(* IEC 61131-3 sources: daoli-st-library/DL_Motion (part 15) *)

(* ---- FB_DL_LaserTabWeldTrack.st ---- *)
(*==============================================================================
 * 组件名称 (Component)  : FB_DL_LaserTabWeldTrack
 * 所属子库 (Sublibrary) : DL_Motion
 * 当前版本 (Version)    : 1.0.1
 * 兼容性 (Platform)     : CODESYS 3.5 / TwinCAT 3 / 汇川 InoProShop（纯标准元素，零方言）
 * 功能描述 (Function)   : 极耳激光焊跟随误差与虚焊特征窗监视。出光期间统计三类缺陷特征
 *                         ——跟随误差超限、功率相对跌落、位置停滞——各需连续满足确认时长
 *                         才置位；单焊点窗口超时强制给出判决并置超时位，绝不允许无限期停
 *                         在出光态。不做激光功率闭环、不做焊缝跟踪插补、不做焊后强度判定。
 *                         交付门槛：位置停滞判据用 tConfirm 换算秒（时间转换链），须在
 *                         CODESYS / TwinCAT / InoProShop 三平台各编译验证一次。
 * 溯源 (Origin)         : 道莅 clean-room 防御性实现
 * 本文件内含 (Contains) : TYPE E_DL_WeldTrackState / FUNCTION_BLOCK FB_DL_LaserTabWeldTrack
 * 依赖 (Depends)        : 无（仅 Standard.library 的 ABS / MAX / TIME_TO_LREAL）
 * 红线自检 (Redline)    : 无外部全局变量、无硬件地址直引 ｜ 全变量中英双语同行注释
 *                         参考功率与误差上限判零防除零 ｜ 位置非有限只跳过本拍、不清峰值
 *                         四个定时器无条件周期刷新 ｜ 枚举显式赋值 ｜ CASE 含 ELSE 兜底
 * 同拍双窗配比约束      : 窗口超时 tWindowMax 必须显著大于三类判据确认 tConfirm
 *                         （建议 tWindowMax ≥ 5 × tConfirm），否则判据来不及确认即被超时
 *                         抢先判决，缺陷掩码永远只能出 bit3。
 * 错误码表 (Codes)      : 16#0004_0331 就绪（无窗进行或本拍无故障）
 *                         16#0004_0332 信息级 位置读数非有限，本拍跳过（已累计峰值与掩码
 *                                    保持，不清零）
 *                         16#0004_0333 故障级 组态非法（跟随误差上限或参考功率 ≤0）
 *                         16#0004_0334 故障级 非法状态兜底（状态机落 ELSE）
 *                         16#0004_0335 预留：本版不发码（下一轮区间起点，禁止回填）
 * 修订历史 (Revision)   : 2026-11-17  v1.0.0  首版入库 · R28 · 阶段三批 2
 *                         2026-11-17  v1.0.1  终审修复：①停滞速度补入组态域闸（负值/NaN 会
 *                                    使停滞距离门限失效而静默关闭 bit2 判据）；②停滞窗起点与
 *                                    焊点位置锁存加位置有限前置（防 NaN 写入出口）· R28 · 阶段四
 * 验收向量 (Acceptance) : 正向 指令 0→50 mm、实际滞后 0.3 mm 超上限 0.2 mm 持续 30 ms →
 *                         bit0 置位、eState=eReject、峰值 0.3 mm
 *                         反向 功率 2000→1500 W（跌 25% 超 10%）持续 30 ms → bit1；
 *                         上限给 0 → 16#0004_0333；窗口拖满 tWindowMax 无判决 → bit3 +
 *                         eReject（不停在出光态）；位置给 NaN → 16#0004_0332 且峰值不清零
 *============================================================================*)

(*-----------------------------------------------------------------------------
 * 枚举: E_DL_WeldTrackState（归属本功能块，同文件发布，全库唯一定义）
 * 含义: 单焊点监视相位，每个成员在 CASE 中有且仅有一个标签。
 *----------------------------------------------------------------------------*)
TYPE E_DL_WeldTrackState :
(
    eWaiting  := 0,    // 待机：等出光 / Waiting for the weld-on signal
    eWelding  := 10,   // 出光中：累计峰值与三类判据 / Welding, accumulating the peak and the three criteria
    eJudging  := 20,   // 判决中：锁存焊点位置并出结论 / Judging, latching the weld position and issuing the verdict
    ePass     := 30,   // 合格：掩码为 0 / Pass, the defect mask is zero
    eReject   := 40,   // 不合格：至少一个缺陷位或窗口超时 / Reject, at least one defect bit or the window timed out
    eFault    := 99    // 故障：锁存码保持，仅使能沿重启 / Fault, the latch code is held until an enable edge
);
END_TYPE

FUNCTION_BLOCK FB_DL_LaserTabWeldTrack
VAR_INPUT
    bEnable         : BOOL := FALSE;      // 使能 / Enable
    bWeldOn         : BOOL := FALSE;      // 出光中（仅窗内判据） / Welding on, the criteria are evaluated inside the window only
    fPosCmd_mm      : REAL := 0.0;        // 指令位置 [mm] / Command position in millimetres
    fPosAct_mm      : REAL := 0.0;        // 实际位置 [mm] / Actual position in millimetres
    fPower_W        : REAL := 0.0;        // 实测功率 [W] / Measured power in watt
    fPowerRef_W     : REAL := 2000.0;     // 设定功率 [W]，须 >0 / Reference power in watt, must be positive
    fFollowErrMax_mm : REAL := 0.2;       // 跟随误差上限 [mm]，域 0.01~2.0 / Following error limit in millimetres, domain 0.01 to 2.0
    fPowerDropPct   : REAL := 10.0;       // 功率跌落阈 [%]，域 1~50 / Power drop threshold in percent, domain 1 to 50
    fStallVel_mmS   : REAL := 0.2;        // 停滞判据速度 [mm/s]，域 0~5 / Stall speed criterion in millimetres per second, domain 0 to 5
    tConfirm        : TIME := T#30MS;     // 判据确认时长 [ms]，域 20~500 / Criterion confirmation time, domain 20 to 500 ms
    tWindowMax      : TIME := T#2S;       // 单焊点窗口 [ms]，域 50ms~10s / Single weld spot window, domain 50 ms to 10 s
END_VAR
VAR_OUTPUT
    bTrackOk        : BOOL;               // 轨迹合格（判决合格时置位） / Trajectory accepted
    fFollowErrPeak_mm : REAL;             // 窗内跟随误差峰值 [mm] / Peak following error inside the window
    uDefectMask     : WORD;               // 缺陷掩码 bit0 跟超 bit1 功率跌 bit2 停滞 bit3 超时 [bit] / Defect mask
    fWeldPos_mm     : REAL;               // 锁存焊点位置 [mm] / Latched weld position in millimetres
    eState          : E_DL_WeldTrackState; // 监视相位 [—] / Monitoring phase
    eErr            : UDINT;              // 错误码，段位 16#0004_xxxx / Error code in segment 16#0004_xxxx
END_VAR
VAR
    _eState         : E_DL_WeldTrackState := E_DL_WeldTrackState.eWaiting; // 当前相位 / Current phase
    _bInit          : BOOL := FALSE;      // 首扫标志，取非判定 / First-scan flag, tested negated
    _bCfgOk         : BOOL;               // 组态合法标志 / Configuration valid flag
    _bPosOk         : BOOL;               // 位置读数有限标志 / Position readings finite flag
    _bFaultLatch    : BOOL;               // 故障锁存标志 / Fault latch flag
    _uLatchCode     : UDINT;              // 锁存码载体 / Latch code carrier
    _fFollowErr     : REAL;               // 本拍跟随误差 [mm] / Following error of this scan
    _fPeak          : REAL;               // 窗内峰值内部副本 [mm] / Internal peak copy inside the window
    _fDropPct       : REAL;               // 本拍功率跌落百分比 [%] / Power drop of this scan in percent
    _fPosWinStart   : REAL;               // 停滞窗起点位置 [mm] / Position at the start of the stall window
    _fConfirmSec    : REAL := 0.03;       // 确认时长换算秒 [s] / Confirmation time converted to seconds
    _fStallDist     : REAL;               // 停滞判定距离门限 [mm] / Stall distance threshold in millimetres
    _rtrigEnable    : R_TRIG;             // 使能上升沿 / Rising edge of the enable input
    _tonFollow      : TON;                // 跟超确认计时 / Following error confirmation timer
    _tonPower       : TON;                // 功率跌落确认计时 / Power drop confirmation timer
    _tonStall       : TON;                // 停滞确认计时 / Stall confirmation timer
    _tonWindow      : TON;                // 单焊点窗口计时 / Weld spot window timer
END_VAR
VAR CONSTANT
    DL_WT_READY     : UDINT := 16#0004_0331;  // 就绪码 / Ready code
    DL_WT_POS_BAD   : UDINT := 16#0004_0332;  // 信息级位置非有限码 / Info code for non-finite positions
    DL_WT_CFG_BAD   : UDINT := 16#0004_0333;  // 故障级组态非法码 / Fault code for bad configuration
    DL_WT_ILLEGAL   : UDINT := 16#0004_0334;  // 故障级非法状态码 / Fault code for an illegal state
    DL_WT_BIT_FOLLOW : WORD := 16#0001;       // 缺陷位 bit0 跟超 / Defect bit 0, following error
    DL_WT_BIT_POWER  : WORD := 16#0002;       // 缺陷位 bit1 功率跌 / Defect bit 1, power drop
    DL_WT_BIT_STALL  : WORD := 16#0004;       // 缺陷位 bit2 停滞 / Defect bit 2, stall
    DL_WT_BIT_TIME   : WORD := 16#0008;       // 缺陷位 bit3 超时 / Defect bit 3, window timeout
    DL_WT_EPS        : REAL := 1.0E-6;        // 浮点判零容差 [—] / Float zero tolerance
END_VAR

// 段 1｜输出与单拍标志预置（bTrackOk 逐拍重算，掩码与峰值为窗内累计量，不在此清）
bTrackOk := FALSE;                                  // 合格标志预清 / Accepted flag pre-cleared
eErr := 0;                                          // 错误码预清 / Error code pre-cleared

// 段 2｜沿检测无条件周期刷新
_rtrigEnable(CLK := bEnable);                       // 使能沿 / Enable edge

// 段 3｜首扫初始化（判据取非，R19）
IF NOT _bInit THEN
    _eState := E_DL_WeldTrackState.eWaiting;        // 相位待机起步 / Phase starts waiting
    _bInit := TRUE;                                 // 首扫只做一次 / The first scan runs once
END_IF

// 段 4｜组态闸（跟随上限与参考功率判零防除零）
_bCfgOk := NOT ((fFollowErrMax_mm <> fFollowErrMax_mm) OR ((fFollowErrMax_mm - fFollowErrMax_mm) <> (fFollowErrMax_mm - fFollowErrMax_mm)))
        AND (fFollowErrMax_mm > DL_WT_EPS)
        AND NOT ((fPowerRef_W <> fPowerRef_W) OR ((fPowerRef_W - fPowerRef_W) <> (fPowerRef_W - fPowerRef_W)))
        AND (fPowerRef_W > DL_WT_EPS)
        AND (fPowerDropPct >= 1.0) AND (fPowerDropPct <= 50.0)
        AND (fStallVel_mmS >= 0.0) AND (fStallVel_mmS <= 5.0)   // 停滞速度域闸：负值/NaN 会使停滞门限失效而静默关闭 bit2 / Stall speed gate, a negative or NaN value silently disables bit 2
        AND (tConfirm >= T#20MS) AND (tConfirm <= T#500MS)
        AND (tWindowMax >= T#50MS) AND (tWindowMax <= T#10S);
_fConfirmSec := TIME_TO_LREAL(tConfirm) / 1000.0;   // 确认时长换算秒 [s] / Confirmation time in seconds
_fStallDist := fStallVel_mmS * _fConfirmSec;        // 停滞判定距离门限 [mm] / Stall distance threshold

// 段 5｜位置有限闸（非有限只跳过本拍，已累计峰值与掩码一律不清零）
_bPosOk := NOT ((fPosCmd_mm <> fPosCmd_mm) OR ((fPosCmd_mm - fPosCmd_mm) <> (fPosCmd_mm - fPosCmd_mm)))
        AND NOT ((fPosAct_mm <> fPosAct_mm) OR ((fPosAct_mm - fPosAct_mm) <> (fPosAct_mm - fPosAct_mm)));
_fFollowErr := ABS(fPosCmd_mm - fPosAct_mm);        // 本拍跟随误差 [mm] / Following error of this scan

// 段 6｜功率跌落百分比（除数已在段 4 判零）
IF (fPower_W <> fPower_W) OR ((fPower_W - fPower_W) <> (fPower_W - fPower_W)) THEN
    _fDropPct := 0.0;                               // 功率非有限：本拍不判跌落 / Non-finite power, no drop judgement this scan
ELSE
    _fDropPct := ((fPowerRef_W - fPower_W) / fPowerRef_W) * 100.0;   // 跌落百分比 [%] / Power drop in percent
END_IF

// 段 7｜四个定时器无条件周期刷新（严禁置于分支内）
_tonFollow(IN := (_eState = E_DL_WeldTrackState.eWelding) AND _bPosOk AND (_fFollowErr > fFollowErrMax_mm), PT := tConfirm);
_tonPower(IN := (_eState = E_DL_WeldTrackState.eWelding) AND (_fDropPct > fPowerDropPct), PT := tConfirm);
_tonStall(IN := (_eState = E_DL_WeldTrackState.eWelding) AND _bPosOk AND (ABS(fPosAct_mm - _fPosWinStart) < _fStallDist), PT := tConfirm);
_tonWindow(IN := (_eState = E_DL_WeldTrackState.eWelding), PT := tWindowMax);

// 段 8｜使能上升沿：锁存解除路径
IF _rtrigEnable.Q THEN
    _bFaultLatch := FALSE;                          // 锁存解除 / Latch released
    _uLatchCode := 0;                               // 锁存码清 / Latch code cleared
    _eState := E_DL_WeldTrackState.eWaiting;        // 相位回待机 / Phase back to waiting
    uDefectMask := 16#0000;                         // 掩码清 / Defect mask cleared
    _fPeak := 0.0;                                  // 峰值清 [mm] / Peak cleared
    fFollowErrPeak_mm := 0.0;                       // 峰值出口清 [mm] / Peak output cleared
END_IF

// 段 9｜失能闸
IF NOT bEnable THEN
    _eState := E_DL_WeldTrackState.eWaiting;        // 相位回待机 / Phase back to waiting
    eErr := DL_WT_READY;                            // 失能为正常停机 / Disable is a normal stop
END_IF

// 段 10｜监视状态机（ENUM + CASE + ELSE 兜底）
IF bEnable THEN
    CASE _eState OF

        E_DL_WeldTrackState.eWaiting:               // 待机：组态错即锁存，出光沿开窗
            IF NOT _bCfgOk THEN
                eErr := DL_WT_CFG_BAD;              // 故障级：组态非法 / Fault, bad configuration
                _uLatchCode := DL_WT_CFG_BAD;
                _bFaultLatch := TRUE;
                _eState := E_DL_WeldTrackState.eFault;
            ELSIF bWeldOn THEN
                uDefectMask := 16#0000;             // 新焊点掩码清 / New spot, the mask is cleared
                _fPeak := 0.0;                      // 新焊点峰值清 [mm] / New spot, the peak is cleared
                fFollowErrPeak_mm := 0.0;
                IF _bPosOk THEN                     // 位置有限才取窗起点与焊点初值（防 NaN 入出口） / Latch only with finite positions
                    _fPosWinStart := fPosAct_mm;    // 停滞窗起点位置 [mm] / Stall window start position
                    fWeldPos_mm := fPosAct_mm;      // 焊点位置初值 [mm] / Weld position initial value
                END_IF
                _eState := E_DL_WeldTrackState.eWelding;   // 开窗出光 / The window opens
            ELSE
                eErr := DL_WT_READY;                // 就绪码 / Ready code
            END_IF

        E_DL_WeldTrackState.eWelding:               // 出光中：累计峰值 + 三类判据确认
            IF NOT _bPosOk THEN
                eErr := DL_WT_POS_BAD;              // 信息级：位置非有限，本拍跳过 / Info, positions not finite, this scan is skipped
            ELSE
                IF _fFollowErr > _fPeak THEN
                    _fPeak := _fFollowErr;          // 峰值刷新 [mm] / Peak refreshed
                END_IF
            END_IF
            fFollowErrPeak_mm := _fPeak;            // 峰值出口 [mm] / Peak output
            IF _fFollowErr > fFollowErrMax_mm THEN
                IF _tonFollow.Q THEN
                    uDefectMask := uDefectMask OR DL_WT_BIT_FOLLOW;   // bit0 跟超确认 / Following error confirmed
                END_IF
            END_IF
            IF _fDropPct > fPowerDropPct THEN
                IF _tonPower.Q THEN
                    uDefectMask := uDefectMask OR DL_WT_BIT_POWER;    // bit1 功率跌落确认 / Power drop confirmed
                END_IF
            END_IF
            IF ABS(fPosAct_mm - _fPosWinStart) < _fStallDist THEN
                IF _tonStall.Q THEN
                    uDefectMask := uDefectMask OR DL_WT_BIT_STALL;    // bit2 停滞确认 / Stall confirmed
                END_IF
            ELSE
                _fPosWinStart := fPosAct_mm;    // 已移动：重置停滞窗起点 [mm] / Moved, restart the stall window
            END_IF
            IF _tonWindow.Q THEN
                uDefectMask := uDefectMask OR DL_WT_BIT_TIME;         // bit3 窗口超时 / Window timed out
                _eState := E_DL_WeldTrackState.eJudging;              // 强制判决，绝不停在出光态 / Forced verdict, never stuck in welding
            ELSIF NOT bWeldOn THEN
                _eState := E_DL_WeldTrackState.eJudging;              // 出光结束：判决 / Weld finished, judge now
            END_IF

        E_DL_WeldTrackState.eJudging:               // 判决中：锁存焊点位置并出结论
            IF _bPosOk THEN                         // 位置有限才刷新焊点位置，保持上次有效值 / Refresh the latch only with finite positions
                fWeldPos_mm := fPosAct_mm;          // 锁存焊点位置 [mm] / Latch the weld position
            END_IF
            IF uDefectMask = 16#0000 THEN
                bTrackOk := TRUE;                   // 掩码为 0：合格 / A zero mask means pass
                _eState := E_DL_WeldTrackState.ePass;
            ELSE
                _eState := E_DL_WeldTrackState.eReject;   // 有缺陷位：不合格 / At least one defect bit, reject
            END_IF
            eErr := DL_WT_READY;                    // 判决本身无故障码 / The verdict produces no fault code

        E_DL_WeldTrackState.ePass:                  // 合格：保持结论，等出光消失后回待机
            bTrackOk := TRUE;
            IF NOT bWeldOn THEN
                _eState := E_DL_WeldTrackState.eWaiting;
            END_IF

        E_DL_WeldTrackState.eReject:                // 不合格：保持结论，等出光消失后回待机
            bTrackOk := FALSE;
            IF NOT bWeldOn THEN
                _eState := E_DL_WeldTrackState.eWaiting;
            END_IF

        E_DL_WeldTrackState.eFault:                 // 故障：锁存码保持
            eErr := _uLatchCode;                    // 锁存码回放 / Replay the latch code
            IF NOT _bFaultLatch THEN
                _eState := E_DL_WeldTrackState.eWaiting;   // 锁存已由使能沿解除 / The latch was released by the enable edge
            END_IF

        ELSE
            // 非法状态兜底（故障级）
            eErr := DL_WT_ILLEGAL;                  // 故障级：非法相位 / Fault, illegal phase
            _uLatchCode := DL_WT_ILLEGAL;
            _bFaultLatch := TRUE;
            _eState := E_DL_WeldTrackState.eFault;

    END_CASE
END_IF

eState := _eState;                                  // 相位出口镜像 / Phase mirrored to the output pin
END_FUNCTION_BLOCK

(* ---- FB_DL_LineShaftClutch.st ---- *)
(*
  FB_DL_LineShaftClutch  —  线轴电子离合器（相位对齐 / 咬合 / 打滑监视 / 强制脱开）/ Line-shaft electronic clutch
  分类 Category : DL_Motion
  码位 Code     : 16#04_0_A2
  版本 Version  : 1.0.2
  来源 Source   : t2-4-s7-motion — IEC 61131-3 标准语义的道莅防御性实现
  溯源 Origin   : S7 Motion Control 公开语义借鉴（电子离合器 / 相位偏移 / 打滑监视），clean-room 实现，未复制源码行
  功能 Function : 1) 对齐段：按相位误差（从轴位置 − 主轴位置 − fPhaseOffsetDeg，归一化到 ±180°）输出修正速度
                     指令 fTrimVelDegS，供下游电子齿轮/速度环消费，误差进 fAlignTolDeg（本件常量 0.5°）后进咬合；
                  2) 咬合段：按 fEngageRampTime 斜坡把同步权重从 0 升到 1，斜坡溢出（TON.Q）置 bEngaged；
                     脱开权重自进入脱开相的实际权重按斜坡线性回落到 0，禁跳变到满值（R38 返修口径）；
                  3) 咬合期监视相位误差，超 fSlipLimitDeg 持续 tSlipDebounce → bSlipFault 锁存并强制脱开；
                  4) 脱开段：按同一斜坡时间把同步权重降回 0，权重回零才回 eIdle（不留残余同步量）。
  边界 Boundary : ① fEngageRampTime <= 0 或 fSlipLimitDeg <= 0 判组态错置 00A2，状态进 eFault 不投运；
                  ② 两轴任一 bError / 非 bEnabled → 拒绝咬合并置信息级 05A2（不置 bError，故障属主是轴本身）；
                  ③ 主从同轴（同一实例注入两侧）判组态错置 04A2：接口契约无指针恒等比较（R28 禁臆造），
                     本件改用**代理判据**——连续 DL_SAME_CYC 拍内两轴位置与速度差均 < 1E-6 且至少一侧使能，
                     视为同一实例注入（说明见「同轴代理判据」段）；
                  ④ 脱开命令与咬合命令同拍 → 以脱开为安全优先（脱开优先判定在本段最前），并置 02A2；
                  ⑤ 咬合中主轴反转（速度 < 0）判工装条件越界 → 强制脱开并置 03A2（反转咬合会拉断机械）；
                  ⑥ bSlipFault 解除式 = bReset AND 主轴 eState = eStandstill AND 从轴 eState = eStandstill
                     （三条件均由注入轴的 PROPERTY 可读，R28-1 通过；接口无 bStandstill 属性，改用
                     E_DL_AxisState.eStandstill 判等，属契约内等价表达，已在头注释声明）。
  依赖 Depends  : I_DL_MotionAxis / E_DL_AxisState（DL_Motion 既有契约件，零修改，仅注入不实例化）；
                  仅 Standard.library（TON / R_TRIG / ABS / MAX / MIN）
  同拍双窗配比  : tSlipDebounce（打滑去抖窗）与 fEngageRampTime 不同源；配比约束
                  tSlipDebounce <= fEngageRampTime × 1000 ms，避免咬合斜坡未完成就打滑判据成立（R100）

  码表 Error codes（本件格 04_0_A2，子码步进 +0x10）:
    16#0004_00A2 故障级：组态非法（斜坡时间 <= 0 / 打滑门限 <= 0 / 对齐容差 <= 0）
    16#0004_01A2 故障级：打滑故障锁存（相位误差超 fSlipLimitDeg 持续 tSlipDebounce，已强制脱开）
    16#0004_02A2 故障级：咬合与脱开命令同拍冲突（脱开优先执行，本码锁存待复位确认）
    16#0004_03A2 故障级：咬合期主轴反转（工装条件越界，已强制脱开）
    16#0004_04A2 故障级：主从同轴注入（代理判据成立，组态错）
    16#0004_05A2 信息级：拒绝咬合（注入轴故障或未使能，不置 bError）
    16#0004_06A2 信息级：咬合完成（bEngaged 上升拍，不置 bError）
    16#0004_07A2 故障级：状态机落 ELSE 兜底（非法相位 ID）
    16#0004_08A2 信息级：脱开起始权重为 0，单拍收口（R38 返修新增，不置 bError）

  修订历史 Revision :
    2026-11-18  v1.0.0  R37 首版
    2026-11-18  v1.0.2  R38 返修：脱离相权重起始值改为进入脱开相快照按斜坡线性回落（_fW0Diseng），起始权重 0 单拍收口，消除反向驱动风险
  R38 已修复    : R37 终审挂账「脱离相耦合权重起始值取成满值」已按快照回落方案修复（六处置相点全部先快照后置相）
*)

TYPE E_DL_ClutchState :
(
    eIdle        := 0,   // 空闲：同步权重 0，等待咬合命令 / Idle, sync weight zero
    eAligning    := 10,  // 对齐中：相位误差收敛至容差内 / Aligning, phase error inside the tolerance
    eRamping     := 20,  // 咬合斜坡中：同步权重 0→1 / Engage ramp, weight rising from zero to one
    eEngaged     := 30,  // 已咬合：同步权重 1，监视打滑 / Engaged, weight one, slip supervised
    eDisengaging := 40,  // 脱开斜坡中：同步权重 1→0 / Disengage ramp, weight falling to zero
    eFault       := 50   // 故障：锁存待复位（复位且两轴静止）/ Fault, latched until reset with both axes standstill
);
END_TYPE

FUNCTION_BLOCK FB_DL_LineShaftClutch
VAR_INPUT
    bEnable        : BOOL := FALSE;              // 总使能，FALSE 时按脱开处理 / Master enable, a low level disengages
    bReset         : BOOL := FALSE;              // 复位，上升沿清故障锁存（须两轴静止）/ Reset, clears the latch when both axes stand still
    bEngageCmd     : BOOL := FALSE;              // 咬合命令（电平，保持型）/ Engage command, level held by the caller
    bDisengageCmd  : BOOL := FALSE;              // 脱开命令（电平，安全优先）/ Disengage command, safety priority
    fPhaseOffsetDeg : REAL := 0.0;               // 从轴相对主轴的相位偏移 [°]，域 ±360 / Phase offset of the slave relative to the master [deg]
    fEngageRampTime : REAL := 0.5;               // 咬合/脱开斜坡时间 [s]，域 > 0 / Engage and disengage ramp time [s]
    fSlipLimitDeg  : REAL := 2.0;                // 打滑门限（相位误差绝对值）[°]，域 > 0 / Slip limit [deg]
    tSlipDebounce  : TIME := T#200MS;            // 打滑去抖窗 [ms]，域 > 0 / Slip debounce window [ms]
    fSlipReleaseBandDeg : REAL := 0.2;           // 打滑解除带回差 [°]，域 >= 0 / Slip release hysteresis band [deg]
END_VAR
VAR_OUTPUT
    bEngaged       : BOOL;                       // 已咬合标志（同步权重达 1）/ Engaged flag, sync weight reached one
    bSlipFault     : BOOL;                       // 打滑故障锁存出口 / Slip fault latch outlet
    fPhaseErrorDeg : REAL;                       // 归一化相位误差 [°]，域 ±180 / Normalised phase error [deg]
    fTrimVelDegS   : REAL;                       // 对齐修正速度指令 [°/s]，带符号 / Alignment trim velocity command [deg/s]
    fSyncWeight    : REAL;                       // 同步权重 [0~1]，供下游齿轮/速度环 / Sync weight for the downstream gear or velocity loop
    bAxesReady     : BOOL;                       // 两轴就绪（使能且无故障）/ Both axes ready
    bError         : BOOL;                       // 故障标志，派生自锁存 / Fault flag derived from the latch
    nErrId         : UDINT;                      // 事件码，0 = 无事件 / Event code, 0 = no event
    eStateOut      : E_DL_ClutchState;           // 状态出口，段尾单点映射 / State outlet, mapped at the tail
END_VAR
VAR_IN_OUT
    iMasterAxis    : I_DL_MotionAxis;            // 主轴接口引用（由调用方注入，本件不实例化）/ Master axis reference, injected
    iSlaveAxis     : I_DL_MotionAxis;            // 从轴接口引用（由调用方注入，本件不实例化）/ Slave axis reference, injected
END_VAR
VAR
    tonRamp        : TON;                        // 咬合/脱开斜坡计时，每拍无条件调用 / Ramp timer, called unconditionally
    tonSlip        : TON;                        // 打滑去抖计时，每拍无条件调用 / Slip debounce timer, called unconditionally
    tonSame        : TON;                        // 同轴代理判据观察窗，自复位 / Same-instance proxy window, self-resetting
    rtReset        : R_TRIG;                     // 复位上升沿 / Reset rising edge
    rtEngaged      : R_TRIG;                     // 咬合完成上升沿（信息码单拍）/ Engaged rising edge, single-scan info code
    _eState        : E_DL_ClutchState := E_DL_ClutchState.eIdle;  // 内部相位（CASE 唯一写入目标）/ Internal phase, the only CASE target
    _uFault        : UDINT;                      // 故障码锁存 / Latched fault code
    _uInfo         : UDINT;                      // 信息码，每拍重算 / Information code, recomputed per scan
    _bFault        : BOOL;                       // 故障锁存位 / Latched fault bit
    _bParamBad     : BOOL;                       // 组态非法聚合 / Configuration invalid aggregate
    _bCmdConflict  : BOOL;                       // 命令同拍冲突 / Command conflict in one scan
    _bReverse      : BOOL;                       // 咬合期主轴反转 / Master reversal while engaged
    _bSlipNow      : BOOL;                       // 打滑判据实时成立 / Slip criterion present
    _bSameAxis     : BOOL;                       // 同轴代理判据成立 / Same-instance proxy verdict
    _bReady        : BOOL;                       // 两轴就绪 / Both axes ready
    _bEngagedPrev  : BOOL;                       // 上拍 bEngaged 快照 / Previous-scan engaged snapshot
    _fPhaseErr     : REAL;                       // 本拍归一化相位误差 [°] / Phase error this scan [deg]
    _fPhaseErrFilt : REAL;                       // 一阶平滑后的相位误差 [°] / First-order smoothed phase error [deg]
    _fWeight       : REAL;                       // 同步权重保持量 [0~1] / Held sync weight
    _fRampSec      : REAL;                       // 生效斜坡时间秒值 [s]，已钳位 / Effective ramp time [s], clamped
    _fPosA         : REAL;                       // 主轴位置快照（一致性比较用）[°] / Master position snapshot [deg]
    _fPosB         : REAL;                       // 从轴位置快照（一致性比较用）[°] / Slave position snapshot [deg]
    _fVelA         : REAL;                       // 主轴速度快照 [°/s] / Master velocity snapshot [deg/s]
    _fVelB         : REAL;                       // 从轴速度快照 [°/s] / Slave velocity snapshot [deg/s]
    _fDeltaPrev    : REAL;                       // 上拍同步权重增量（脱开斜坡复用）[1] / Previous weight increment, reused by the disengage ramp
    _fW0Diseng     : REAL := 0.0;                // 脱开起始权重快照（进入脱开相当拍的实际权重）/ Snapshot of the weight at the disengage entry
    _bRampBreak    : BOOL := TRUE;               // 斜坡计时断输入一拍（相位入口重启，防沿用上段 ET）/ One-scan ramp break to restart the timer at a phase entry
END_VAR
VAR CONSTANT
    DL_ALIGN_TOL_DEG : REAL := 0.5;      // 对齐容差 [°]，本件声明常量（规格固定值）/ Alignment tolerance, fixed by the specification
    DL_ALIGN_KP      : REAL := 2.0;      // 对齐比例增益 [1/s] / Alignment proportional gain
    DL_TRIM_MAX_DEGS : REAL := 90.0;     // 修正速度饱和上限 [°/s] / Trim velocity saturation limit
    DL_RAMP_MAX_SEC  : REAL := 60.0;     // 斜坡时间上限 [s] / Ramp time ceiling
    DL_EPS           : REAL := 1.0E-6;   // 判零容差 [1] / Zero tolerance
    DL_SAME_CYC      : TIME := T#2S;     // 同轴观察窗 [ms]，自复位节拍 / Same-instance window, self-resetting
    DL_POS_WRAP      : REAL := 360.0;    // 位置一圈对应角度 [°] / One full revolution in degrees
    DL_POS_HALF      : REAL := 180.0;    // 归一化半圈 [°] / Half revolution used by the normalisation
    DL_FILT_ALPHA    : REAL := 0.35;     // 相位误差一阶平滑系数 [1] / Phase error smoothing coefficient
    DL_W0_EPS        : REAL := 1.0E-6;   // 脱开起始权重判零阈 [1]（R38 返修新增）/ Zero threshold for the disengage entry weight
END_VAR

(* —— 段 0：定时器与边缘检测无条件周期刷新（R182：禁置于 IF / CASE 内） —— *)
rtReset(CLK := bReset);                                          // 复位上升沿，每拍必调
rtEngaged(CLK := bEngaged);                                      // 咬合完成上升沿，每拍必调
tonSame(IN := NOT tonSame.Q, PT := DL_SAME_CYC);                 // 同轴观察窗自复位：到点下一拍断输入
tonRamp(IN := (((_eState = E_DL_ClutchState.eRamping) OR (_eState = E_DL_ClutchState.eDisengaging))
               AND (NOT _bRampBreak)),
        PT := REAL_TO_TIME(_fRampSec * 1000.0));                  // 斜坡计时（条件以表达式传入，调用本身无条件）
_bRampBreak := FALSE;                                             // 断输入拍在调用后自清（相位入口置位）
tonSlip(IN := (_eState = E_DL_ClutchState.eEngaged) AND _bSlipNow,
        PT := tSlipDebounce);                                     // 打滑去抖计时（表达式入参，调用无条件）

(* —— 段 1：单拍量预清零（快照 / 锁存 / 权重不入清单，R187①） —— *)
_uInfo        := 16#0000_0000;   // 信息码每拍重算
bError        := FALSE;          // 故障出口每拍重算，段 7 由锁存派生
bEngaged      := FALSE;          // 咬合出口缺省 FALSE，段 6 单点置位
bAxesReady    := FALSE;          // 就绪出口缺省 FALSE
_bParamBad    := FALSE;          // 组态非法预清零
_bCmdConflict := FALSE;          // 命令冲突预清零
_bReverse     := FALSE;          // 反转标志预清零
_bSameAxis    := FALSE;          // 同轴代理标志预清零

(* —— 段 2：复位沿清锁存（打滑故障解除式含两轴静止条件，R28-1） —— *)
IF rtReset.Q THEN
    IF (iMasterAxis.eState = E_DL_AxisState.eStandstill) AND
       (iSlaveAxis.eState = E_DL_AxisState.eStandstill) THEN
        _bFault := FALSE;            // 两轴静止：解除打滑/冲突/反转类锁存
        _uFault := 16#0000_0000;     // 锁存码同拍清除
    END_IF
END_IF

(* —— 段 3：组态域闸（覆盖全部参与换算的引脚，R151） —— *)
_fRampSec := fEngageRampTime;                       // 斜坡时间直取引脚 [s]
IF (_fRampSec <> _fRampSec) OR (_fRampSec <= 0.0) THEN
    _bParamBad := TRUE;                             // 斜坡时间非法（权重增量的分母）
END_IF
IF _fRampSec > DL_RAMP_MAX_SEC THEN
    _fRampSec := DL_RAMP_MAX_SEC;                   // 上限钳位（防权重增量下溢为 0）
END_IF
IF (fSlipLimitDeg <> fSlipLimitDeg) OR (fSlipLimitDeg <= 0.0) THEN
    _bParamBad := TRUE;                             // 打滑门限非法
END_IF
IF (fSlipReleaseBandDeg <> fSlipReleaseBandDeg) OR (fSlipReleaseBandDeg < 0.0) THEN
    _bParamBad := TRUE;                             // 解除回差非法（负值会让判据自相矛盾）
END_IF
IF (fPhaseOffsetDeg <> fPhaseOffsetDeg) OR (ABS(fPhaseOffsetDeg) > DL_POS_WRAP) THEN
    _bParamBad := TRUE;                             // 相位偏移非法（超一圈无物理意义）
END_IF
IF _bParamBad THEN
    _uFault := 16#0004_00A2;                        // 故障级：组态非法
    _bFault := TRUE;                                // 锁存位置位（复位沿可清）
    bError  := TRUE;                                // 故障标志置位（R45 配对）
    _eState := E_DL_ClutchState.eFault;             // 状态机进故障相
END_IF

(* —— 段 4：轴状态采集与同轴代理判据（只读接口属性，零命令下发） —— *)
_fPosA := iMasterAxis.fPosition;                    // 主轴位置 [°]
_fPosB := iSlaveAxis.fPosition;                     // 从轴位置 [°]
_fVelA := iMasterAxis.fVelocity;                    // 主轴速度 [°/s]
_fVelB := iSlaveAxis.fVelocity;                     // 从轴速度 [°/s]
_bReady := iMasterAxis.bEnabled AND iSlaveAxis.bEnabled AND
           (NOT iMasterAxis.bError) AND (NOT iSlaveAxis.bError);   // 两轴就绪（接口契约仅提供 bError，无 bFault 属性）
bAxesReady := _bReady;                              // 就绪出口（诊断用，不影响状态迁移）

IF (ABS(_fPosA - _fPosB) < DL_EPS) AND (ABS(_fVelA - _fVelB) < DL_EPS) AND
   (iMasterAxis.bEnabled OR iSlaveAxis.bEnabled) THEN
    IF tonSame.Q THEN
        _bSameAxis := TRUE;                         // 持续一整窗完全重合：代理判据成立（同一实例注入）
    END_IF
END_IF
IF _bSameAxis THEN
    _uFault := 16#0004_04A2;                        // 故障级：主从同轴注入（组态错）
    _bFault := TRUE;                                // 锁存
    bError  := TRUE;                                // 故障标志置位（R45 配对）
    _eState := E_DL_ClutchState.eFault;             // 进故障相
END_IF

(* —— 段 5：相位误差与打滑判据（无故障时计算，故障期保持末值） —— *)
IF NOT _bFault THEN
    _fPhaseErr := _fPosB - _fPosA - fPhaseOffsetDeg;            // 原始相位误差 [°]
    IF _fPhaseErr > DL_POS_HALF THEN
        _fPhaseErr := _fPhaseErr - DL_POS_WRAP;                 // 归一化：超 +180 折回负半圈 [°]
    END_IF
    IF _fPhaseErr < -DL_POS_HALF THEN
        _fPhaseErr := _fPhaseErr + DL_POS_WRAP;                 // 归一化：低于 −180 折回正半圈 [°]
    END_IF
    _fPhaseErrFilt := _fPhaseErrFilt + DL_FILT_ALPHA * (_fPhaseErr - _fPhaseErrFilt);  // 一阶平滑（抗单点毛刺）
    fPhaseErrorDeg := _fPhaseErrFilt;                           // 出口取平滑值
    _bSlipNow := (ABS(_fPhaseErrFilt) > fSlipLimitDeg);         // 打滑判据（实时）
    IF (_eState = E_DL_ClutchState.eEngaged) AND (_fVelA < -DL_EPS) THEN
        _bReverse := TRUE;                                      // 咬合期主轴反转：工装条件越界
    END_IF
    IF bDisengageCmd AND bEngageCmd THEN
        _bCmdConflict := TRUE;                                  // 同拍冲突：脱开优先（安全优先）
    END_IF
END_IF

(* —— 段 6：相位机（只做迁移与权重演进；输出映射在段 8） —— *)
CASE _eState OF

E_DL_ClutchState.eIdle:
    _fWeight := 0.0;                                            // 空闲：同步权重归零（唯一清零点在本相）
    IF bDisengageCmd THEN
        _fW0Diseng := _fWeight;                                 // R38 返修：空闲拍脱开命令 sighted，快照保持新鲜（本相权重恒 0）
        _uInfo := 16#0004_05A2;                                 // 空闲拍收到脱开：无需动作（信息级，不置错）
    ELSIF bEngageCmd THEN
        IF (NOT _bReady) THEN
            _uInfo := 16#0004_05A2;                             // 拒绝咬合：轴故障或未使能（信息级）
        ELSIF _bCmdConflict THEN
            _uFault := 16#0004_02A2;                            // 故障级：命令同拍冲突，脱开优先
            _bFault := TRUE;                                    // 锁存
            bError  := TRUE;                                    // 故障标志置位（R45 配对）
            _eState := E_DL_ClutchState.eFault;                 // 进故障相
        ELSE
            _eState := E_DL_ClutchState.eAligning;              // 进对齐相
            _fPhaseErrFilt := _fPhaseErr;                       // 平滑器赋初值，防首拍冲击
        END_IF
    END_IF

E_DL_ClutchState.eAligning:
    IF bDisengageCmd OR (NOT bEnable) THEN
        _fW0Diseng := _fWeight;                                 // R38 返修：先快照进入脱开相的实际权重（本相恒 0）
        _eState := E_DL_ClutchState.eDisengaging;               // 脱开命令/失能：回脱开斜坡（权重快照 0，单拍收口）
        _bRampBreak := TRUE;                                    // 脱开斜坡计时从零重启
    ELSIF NOT _bReady THEN
        _uInfo := 16#0004_05A2;                                 // 轴掉就绪：退出对齐（信息级，不置错）
        _eState := E_DL_ClutchState.eIdle;
    ELSIF ABS(_fPhaseErrFilt) <= DL_ALIGN_TOL_DEG THEN
        _eState := E_DL_ClutchState.eRamping;                   // 误差进容差：进咬合斜坡
        _fWeight := 0.0;                                        // 斜坡起点权重归零（迁移拍归零，非同拍抹除）
        _bRampBreak := TRUE;                                    // 斜坡计时从零重启，不沿用对齐段残留
    END_IF

E_DL_ClutchState.eRamping:
    (* 本相权重由段 6A 按 TON.ET 比例推进，此处不写 _fWeight，避免双写同拍覆盖 *)
    IF bDisengageCmd OR (NOT bEnable) THEN
        _fW0Diseng := _fWeight;                                 // R38 返修：先快照斜坡中途的实际权重（0~1 区间）
        _eState := E_DL_ClutchState.eDisengaging;               // 脱开优先
        _bRampBreak := TRUE;                                    // 脱开斜坡计时从零重启（不沿用咬合段 ET）
    ELSIF NOT _bReady THEN
        _fW0Diseng := _fWeight;                                 // R38 返修：轴掉就绪路径同样先快照
        _eState := E_DL_ClutchState.eDisengaging;               // 轴掉就绪：按脱开处理（不锁存故障）
        _bRampBreak := TRUE;                                    // 脱开斜坡计时从零重启
    ELSIF ABS(_fPhaseErrFilt) > fSlipLimitDeg THEN
        _uFault := 16#0004_01A2;                                // 斜坡期越打滑门限：直接判打滑（斜坡未完成不得掩盖）
        _bFault := TRUE;                                        // 锁存
        bError  := TRUE;                                        // 故障标志置位（R45 配对）
        _eState := E_DL_ClutchState.eFault;                     // 进故障相
    ELSIF tonRamp.Q THEN
        _eState := E_DL_ClutchState.eEngaged;                   // 斜坡完成：已咬合
        _fWeight := 1.0;                                        // 权重锁定为 1
        _uInfo := 16#0004_06A2;                                 // 信息级：咬合完成
    END_IF

E_DL_ClutchState.eEngaged:
    _fWeight := 1.0;                                            // 已咬合：权重保持 1
    IF bDisengageCmd OR (NOT bEnable) THEN
        _fW0Diseng := _fWeight;                                 // R38 返修：已咬合（权重 1）正常脱开先快照
        _eState := E_DL_ClutchState.eDisengaging;               // 正常脱开
        _bRampBreak := TRUE;                                    // 脱开斜坡计时从零重启
    ELSIF NOT _bReady THEN
        _fW0Diseng := _fWeight;                                 // R38 返修：轴掉就绪路径先快照（权重 1）
        _eState := E_DL_ClutchState.eDisengaging;               // 轴掉就绪：脱开但不锁存（故障属主为轴）
        _bRampBreak := TRUE;                                    // 脱开斜坡计时从零重启
    ELSIF _bReverse THEN
        _uFault := 16#0004_03A2;                                // 故障级：咬合期主轴反转
        _bFault := TRUE;                                        // 锁存
        bError  := TRUE;                                        // 故障标志置位（R45 配对）
        _eState := E_DL_ClutchState.eFault;                     // 强制脱开（进故障相即权重归零）
    ELSIF tonSlip.Q THEN
        _uFault := 16#0004_01A2;                                // 故障级：打滑故障锁存
        _bFault := TRUE;                                        // 锁存
        bError  := TRUE;                                        // 故障标志置位（R45 配对）
        _eState := E_DL_ClutchState.eFault;                     // 强制脱开
    END_IF

E_DL_ClutchState.eDisengaging:
    IF _fW0Diseng <= DL_W0_EPS THEN
        _fWeight := 0.0;                                        // R38 返修：起始权重为 0 → 不等斜坡单拍收口（兑现原注释语义）
        _eState := E_DL_ClutchState.eIdle;                      // 直回空闲
        _uInfo := 16#0004_08A2;                                 // 信息级：脱开起始权重为 0，单拍收口
    ELSIF tonRamp.Q THEN
        _fWeight := 0.0;                                        // 斜坡到点：权重归零（脱开完成）
        _eState := E_DL_ClutchState.eIdle;                      // 回空闲
    END_IF

E_DL_ClutchState.eFault:
    _fWeight := 0.0;                                            // 故障：同步权重强制 0（机械不再被拖动）
    IF (NOT _bFault) THEN
        _eState := E_DL_ClutchState.eIdle;                      // 锁存已由复位沿清除：回空闲重新对齐
    END_IF

ELSE
    _uFault := 16#0004_07A2;                                    // 故障级：相位 ID 越界（枚举兜底）
    _bFault := TRUE;                                            // 锁存
    bError  := TRUE;                                            // 故障标志置位（R45 配对）
    _eState := E_DL_ClutchState.eFault;                         // 强制回故障相
END_CASE

(* —— 段 6A：权重演进（唯一累加点；脱开斜坡按 TON 比例回落，禁在 CASE 内二次写） —— *)
IF _eState = E_DL_ClutchState.eRamping THEN
    _fWeight := MIN(1.0, TIME_TO_REAL(tonRamp.ET) / (_fRampSec * 1000.0));  // 咬合权重按斜坡比例上升（分母已证 > 0）
ELSIF _eState = E_DL_ClutchState.eDisengaging THEN
    _fWeight := MAX(0.0, _fW0Diseng * (1.0 - TIME_TO_REAL(tonRamp.ET) / (_fRampSec * 1000.0)));  // R38 返修：按进入脱开相的快照权重线性回落到 0，禁跳变到满值
END_IF

(* —— 段 7：对齐修正速度与故障码优先级链（每个 bError 置位源均在此有码，R45） —— *)
IF _eState = E_DL_ClutchState.eAligning THEN
    fTrimVelDegS := _fPhaseErrFilt * DL_ALIGN_KP;               // 比例修正速度 [°/s]
    IF fTrimVelDegS > DL_TRIM_MAX_DEGS THEN
        fTrimVelDegS := DL_TRIM_MAX_DEGS;                       // 上行饱和（防超速）
    END_IF
    IF fTrimVelDegS < -DL_TRIM_MAX_DEGS THEN
        fTrimVelDegS := -DL_TRIM_MAX_DEGS;                      // 下行饱和
    END_IF
ELSE
    fTrimVelDegS := 0.0;                                        // 非对齐相：修正速度 0（语义：不对轴施加修正）
END_IF

(* —— 段 8：出口单点映射（名实同源；锁存码回放，禁同拍抹除） —— *)
bEngaged     := (_eState = E_DL_ClutchState.eEngaged);          // 咬合出口：仅 eEngaged 相为真
bSlipFault   := _bFault AND (_uFault = 16#0004_01A2);           // 打滑故障出口：按码定向，不与其它锁存混用
fSyncWeight  := _fWeight;                                       // 同步权重出口
eStateOut    := _eState;                                        // 状态出口
IF _bFault THEN
    nErrId := _uFault;                                          // 故障锁存码回放（不在故障相按当下输入重推）
    bError := TRUE;                                             // 故障出口派生自锁存
ELSE
    nErrId := _uInfo;                                           // 信息码
END_IF

END_FUNCTION_BLOCK

(* ---- FB_DL_LoadShareDroop.st ---- *)
(*==============================================================================
 * 组件名称 (Component)  : FB_DL_LoadShareDroop
 * 所属子库 (Sublibrary) : DL_Motion
 * 当前版本 (Version)    : 1.0.0
 * 兼容性   (Platform)   : CODESYS 3.5+ / TwinCAT 3 / 汇川 InoProShop / 施耐德 Machine Expert
 *                         仅依赖 Standard.library（ABS / MIN / MAX），零厂商私有库
 * 功能描述 (Function)   : 多轴（≤4）负载均衡 droop 调差：按各轴负载百分比对速度基准做
 *                         droop 修正，负载高于均值者减速让载、低于均值者提速分担：
 *                           aVout[i] = fVref × (1 - fDroopPct × (aLoad[i]-fLoadAvg)/100)
 *                         均衡目标带内（|aLoad[i]-fLoadAvg| <= fShareBandPct）不修正
 *                         （死区防振荡）；非负载轴（bAxActive=FALSE）输出直通不修正；
 *                         均值只对有效轴计算。
 * 接口     (Interface)  : 输入 fVrefMmS 速度基准（mm/s）、aLoadPct 各轴负载（%，定长
 *                         1..nAxMax 数组）、bAxActive 各轴有效、fDroopPct 调差率
 *                         （%/(100%负载)）、fShareBandPct 均衡目标带（%）、fVrefMax 输出
 *                         钳限（mm/s）；输出 aVoutMmS 各轴修正后速度（mm/s）、bBalanced
 *                         均衡达标、bNoLoad 全轴失效。
 * 边界     (Boundary)   : ① **属主边界（写死）：本件只做速度基准的 droop 修正分配，不写
 *                         轴指令、不接管同步耦合**；几何同步归 `FB_DL_GantrySyncAxis`，
 *                         偏差监视归 `FB_DL_GantrySkewMonitor`（修调 ≠ 监视）。
 *                         ② 数组边界逐轴钳位（索引 1..nAxMax 常量域，循环定界，无越界路径）。
 *                         ③ 全轴失效（无有效轴）→ 直通输出 fVref 并置 bNoLoad（均值除零
 *                         前置：有效轴计数 >= 1 才算均值，R28 防除零）。
 *                         ④ 非有限负载当拍该轴按失效处理（不入均值、输出直通）并置当拍
 *                         bError（R245）；fVref 非有限 → 全轴直通冻结。
 *                         ⑤ 输出钳 ±fVrefMax（fVrefMax 组态域闸 > 0，锁存 bError，
 *                         解除沿 = 无（无复位引脚，组态合法化后自动解除，头注释声明：
 *                         组态闸为当拍判据非锁存，修正组态即解除）。
 *                         ⑥ 零全局耦合（无 GVL / VAR_EXTERNAL / 物理地址）。
 * 分工声明 (Scope)      : 与 `FB_DL_GantrySyncAxis` 分工：负载均衡 ≠ 几何同步；与
 *                         `FB_DL_GantrySkewMonitor` 分工：修调 ≠ 监视。
 * 来源标签 (Source Tag) : T1-6 ◐（PLCopen MC 语义只借多轴协同语义，droop 公式为电力
 *                         系统公开调差定义 clean-room）
 * 码表     (Codes)      : 本件不占用任何全局数字码位。出口为 LREAL 数组 + BOOL 组；
 *                         数字码位待主控收口阶段统一派号。
 * 红线自检 (Redline)    : R1 ✓ 零 GVL/VAR_EXTERNAL ｜ R2 ✓ 零 %I/%Q/%M ｜ R3 ✓ 纯 IEC 61131-3
 *                         R4 ✓ 均值除零前置 + 非有限剔除 + 输出钳位 ｜ R5 ✓ 声明逐行同行双语注释
 *                         R6 N/A（无状态机） ｜ R7 N/A（无实例调用）
 * 修订历史 (Revision)   : 2026-11-20  v1.0.0  R48 首版（批次 3 · 序号 14）
 *                         验收向量：双轴等载 → 无修正；单轴 120% 均值 → 该轴减速；
 *                         全轴失效 → 直通 + bNoLoad；带内不修正防振荡。
 *==============================================================================*)

FUNCTION_BLOCK FB_DL_LoadShareDroop
VAR_INPUT
    fVrefMmS     : LREAL := 100.0;                       // 速度基准 [mm/s] / Velocity reference [mm/s]
    aLoadPct     : ARRAY[1..4] OF LREAL := [0.0, 0.0, 0.0, 0.0];   // 各轴负载（0~100+） [%] / Per-axis load [%]
    bAxActive    : ARRAY[1..4] OF BOOL := [FALSE, FALSE, FALSE, FALSE];   // 各轴参与均衡有效标志 [-] / Per-axis active flag
    fDroopPct    : LREAL := 5.0;                         // 调差率（每 100% 负载偏差的速度降幅） [%/(100%负载)] / Droop rate
    fShareBandPct: LREAL := 2.0;                         // 均衡目标带半宽（带内不修正） [%] / Balance target band [%]
    fVrefMax     : LREAL := 150.0;                       // 输出钳限（对称 ±），域 > 0 [mm/s] / Output clamp limit [mm/s]
END_VAR
VAR_OUTPUT
    aVoutMmS  : ARRAY[1..4] OF LREAL;                    // 各轴修正后速度输出 [mm/s] / Per-axis corrected velocity output
    bBalanced : BOOL;                                    // 均衡达标（全部有效轴在目标带内） [-] / Balanced flag
    bNoLoad   : BOOL;                                    // 全轴失效直通标志 [-] / No active axis flag
    bError    : BOOL;                                    // 故障标志（组态病 ∨ 输入病当拍） [-] / Error flag
END_VAR
VAR
    _nActive  : DINT;            // 有效轴计数 [轴] / Active axis count
    _fSum     : LREAL;           // 有效轴负载和 [%] / Active load sum
    _fAvg     : LREAL;           // 有效轴负载均值 [%] / Active load mean
    _fDev     : LREAL;           // 单轴负载对均值偏差 [%] / Per-axis load deviation
    _fOut     : LREAL;           // 单轴修正中间量 [mm/s] / Per-axis corrected intermediate
    _bBal     : BOOL;            // 均衡达标内部量 / Balanced internal
    _bErrScan : BOOL;            // 输入病当拍量 [-] / Per-scan input fault
    _bCfgBad  : BOOL;            // 组态病当拍量（fVrefMax<=0，当拍判据非锁存） / Config fault this scan
    i         : DINT;            // 轴循环索引（1..4 定界） / Axis loop index
END_VAR
VAR CONSTANT
    DL_LSD_NAX  : DINT  := 4;        // 支持轴数上限（数组定界） [轴] / Supported axis ceiling
    DL_LSD_PCT  : LREAL := 100.0;    // 百分比换算基 [无量纲] / Percent conversion base
    DL_LSD_EPS  : LREAL := 0.0;      // 非有限差值判零基准 [-] / Non-finite difference zero base
END_VAR

(* —— 段 0：组态闸 + 输入病判（当拍判据，非锁存，头注释⑤声明解除语义） —— *)
_bCfgBad := fVrefMax <= 0.0;                                 // 钳限组态闸 / Clamp config gate
_bErrScan := (fVrefMmS <> fVrefMmS) OR ((fVrefMmS - fVrefMmS) <> DL_LSD_EPS);   // 基准非有限（R245） / Non-finite reference
FOR i := 1 TO DL_LSD_NAX DO
    IF bAxActive[i] AND ((aLoadPct[i] <> aLoadPct[i]) OR ((aLoadPct[i] - aLoadPct[i]) <> DL_LSD_EPS)) THEN
        _bErrScan := TRUE;                                   // 有效轴负载非有限：当拍输入病（R245） / Non-finite load on active axis
    END_IF
END_FOR

(* —— 段 1：直通总闸（组态病 ∨ 基准非有限 → 全轴直通） —— *)
bNoLoad := FALSE;                                            // 全轴失效标志预清 / No-load preset
IF _bCfgBad OR _bErrScan THEN
    FOR i := 1 TO DL_LSD_NAX DO
        aVoutMmS[i] := fVrefMmS;                             // 全轴直通基准（直通即语义，头注释④） / Pass-through all axes
    END_FOR
    bBalanced := FALSE;                                      // 直通期不报均衡达标 / Not balanced
ELSE
    (* 段 2：有效轴均值（计数 >= 1 才除，无除零） *)
    _nActive := 0;                                           // 有效计数清零 / Clear count
    _fSum := 0.0;                                            // 负载和清零 / Clear sum
    FOR i := 1 TO DL_LSD_NAX DO
        IF bAxActive[i] THEN
            _nActive := _nActive + 1;                        // 有效轴计数 / Count active axis
            _fSum := _fSum + aLoadPct[i];                    // 累加有效负载 / Accumulate load
        END_IF
    END_FOR
    IF _nActive >= 1 THEN
        _fAvg := _fSum / DINT_TO_LREAL(_nActive);            // 有效轴均值（分母计数已闸） / Active mean
        _bBal := TRUE;                                       // 均衡达标预置（任一越带即翻假） / Balanced preset
        FOR i := 1 TO DL_LSD_NAX DO
            IF bAxActive[i] THEN
                _fDev := aLoadPct[i] - _fAvg;                // 负载对均值偏差 [%] / Load deviation
                IF ABS(_fDev) <= fShareBandPct THEN
                    aVoutMmS[i] := fVrefMmS;                 // 带内不修正（死区防振荡） / In-band: no correction
                ELSE
                    _fOut := fVrefMmS * (1.0 - fDroopPct * _fDev / DL_LSD_PCT);   // droop 调差修正（高载减速让载） / Droop correction
                    IF _fOut > fVrefMax THEN
                        _fOut := fVrefMax;                   // 输出上钳 ±fVrefMax / Clamp high
                    ELSIF _fOut < -fVrefMax THEN
                        _fOut := -fVrefMax;                  // 输出下钳 / Clamp low
                    END_IF
                    aVoutMmS[i] := _fOut;                    // 修正输出 / Corrected output
                    _bBal := FALSE;                          // 有轴越带：未均衡 / Axis out of band
                END_IF
            ELSE
                aVoutMmS[i] := fVrefMmS;                     // 非负载轴直通不修正（头注释①） / Inactive axis pass-through
            END_IF
        END_FOR
        bNoLoad := FALSE;                                    // 有有效轴 / Load exists
        bBalanced := _bBal;                                  // 均衡达标出口 / Balanced outlet
    ELSE
        FOR i := 1 TO DL_LSD_NAX DO
            aVoutMmS[i] := fVrefMmS;                         // 全轴失效：直通（均值除零前置跳过） / No active axis: pass-through
        END_FOR
        bNoLoad := TRUE;                                     // 置全轴失效标志 / Raise no-load flag
        bBalanced := FALSE;                                  // 无轴谈不上均衡 / Not balanced
    END_IF
END_IF

(* —— 段 3：故障出口（组态病 ∨ 输入病，R191 同源） —— *)
bError := _bCfgBad OR _bErrScan;                             // 故障标志出口 / Error flag outlet

END_FUNCTION_BLOCK

(* ---- FB_DL_LookaheadVelPlanner.st ---- *)
(*==============================================================================
 * 组件名称 (Component)  : FB_DL_LookaheadVelPlanner
 * 所属子库 (Sublibrary) : DL_Motion
 * 当前版本 (Version)    : 1.0.1
 * 兼容性   (Platform)   : CODESYS 3.5+ / TwinCAT 3 / 汇川 InoProShop / 施耐德 Machine Expert
 *                         仅依赖 Standard.library（MIN / SQRT），零厂商私有库
 * 功能描述 (Function)   : 多段路径前瞻速度规划（回溯-前传两遍法）：输入段几何表（段长 /
 *                         拐角半径 / 段限速 / 段加速度）与轨迹目标速度，输出各段允许速度
 *                         上限表，供段执行器逐段限速。三步：
 *                         ① 拐角限速 fVcorner = SQRT(fAccel × fCornerRad)（向心加速度
 *                            <= fAccel 推导式，段直通无拐角时 fCornerRad=0 → 0 不限）；
 *                         ② 自深至浅回溯（减速可达性反推，前瞻深度 nLookahead）：
 *                            aVelCap[i]² = MIN(aVelCap[i]², aVelCap[i+1]² + 2×fAccel[i]
 *                            × fLen[i+1])（累加式为负先钳 0 再开方）；
 *                         ③ 前向传播可达上限：aVelCap[i+1]² = MIN(aVelCap[i+1]²,
 *                            aVelCap[i]² + 2×fAccel[i+1] × fLen[i+1])。
 * 接口     (Interface)  : 输入 aSeg 段几何表（定长 1..nSegMax）、nSegCount 有效段数、
 *                         nLookahead 前瞻深度、fVtrajMmS 轨迹目标速度（mm/s）、bReset
 *                         复位；输出 aVelCapMmS 各段速度上限（mm/s）、bPlanned 规划完成
 *                         单拍、bCfgBad 组态非法（锁存）、bError 故障标志。
 * 边界     (Boundary)   : ① **属主边界（写死）：本件只出段速度上限表，不生成速度曲线、
 *                         不排队指令**（单段成形归 `FB_DL_SCurveGenerator`，指令排队归
 *                         `FB_DL_MotionCmdQueue`）。
 *                         ② nSegCount=0 或超 nSegMax 钳位并报组态（锁存 bCfgBad）。
 *                         ③ 段几何病：fLen<=0 / fAccel<=0 / fVmax<=0 → 锁存 bCfgBad
 *                         （零长度段除零隐患前置，规格边界）；病态期输出冻结。
 *                         ④ SQRT 前判负：回溯累加式 aVelCap[i+1]² + 2×a×L 可能为负，
 *                         先钳 0 再开方（规格边界）。
 *                         ⑤ 回溯/前传用 FOR 定界循环（界宽 = nLookahead 与 nSegCount 钳位
 *                         后的最小值，迭代次数静态有界，等价 WHILE+步数计数防死锁且无
 *                         死锁可能，头注释声明实现选择）。
 *                         ⑥ 零全局耦合（无 GVL / VAR_EXTERNAL / 物理地址）。
 * 分工声明 (Scope)      : 与 `FB_DL_SCurveGenerator` 分工：段间衔接规划 ≠ 单段 S 曲线
 *                         成形；与 `FB_DL_MotionCmdQueue` 分工：几何规划 ≠ 指令排队。
 * 来源标签 (Source Tag) : T1-6 ◐（PLCopen MC 语义只借前瞻规划语义，回溯-前传两遍法为
 *                         公开规划算法 clean-room）
 * 码表     (Codes)      : 本件不占用任何全局数字码位。出口为 LREAL 数组 + BOOL 组；
 *                         数字码位待主控收口阶段统一派号。
 * 红线自检 (Redline)    : R1 ✓ 零 GVL/VAR_EXTERNAL ｜ R2 ✓ 零 %I/%Q/%M ｜ R3 ✓ 纯 IEC 61131-3
 *                         R4 ✓ 段病锁存 + SQRT 前钳负 + 计数钳位 ｜ R5 ✓ 声明逐行同行双语注释
 *                         R6 N/A（规划无状态机） ｜ R7 ✓ 一 R_TRIG 段 0 无条件刷新
 * 修订历史 (Revision)   : 2026-11-20  v1.0.1  R50 返修 R1：回溯步减速距离误用
 *                         邻段长度 L[i+1]，更正为本段 L[i]（与前传步取
 *                         L[i+1] 前后对称一致）；行为变更同步更新验收向量。
 *                         2026-11-20  v1.0.0  R48 首版（批次 4 · 序号 17）
 *                         验收向量：三段直角路径回溯降速；拐角半径 0 段不限；前瞻深度
 *                         截断；零长度段 → bCfgBad 锁存。
 *==============================================================================*)

TYPE ST_DL_SegGeom :
STRUCT
    fLenMm    : LREAL;   // 段长度，域 > 0 [mm] / Segment length [mm]
    fCornerRad: LREAL;   // 段末拐角半径（0=直通无限速） [mm] / Corner radius at segment end [mm]
    fVmaxMmS  : LREAL;   // 段自身限速，域 > 0 [mm/s] / Segment speed ceiling [mm/s]
    fAccelMmS2: LREAL;   // 段加减速度能力，域 > 0 [mm/s²] / Segment acceleration capability [mm/s2]
END_STRUCT
END_TYPE

FUNCTION_BLOCK FB_DL_LookaheadVelPlanner
VAR_INPUT
    aSeg      : ARRAY[1..16] OF ST_DL_SegGeom;   // 段几何表（定长，nSegCount 指明有效前段） / Segment geometry table
    nSegCount : UDINT := 0;     // 有效段数（0=组态非法） [段] / Valid segment count
    nLookahead: UDINT := 4;     // 前瞻深度（回溯跨越的段数） [段] / Lookahead depth in segments
    fVtrajMmS : LREAL := 200.0; // 轨迹目标速度，域 > 0 [mm/s] / Trajectory target speed [mm/s]
    bReset    : BOOL := FALSE;  // 复位，上升沿清 bCfgBad 锁存 [-] / Reset, rising edge clears cfg latch
END_VAR
VAR_OUTPUT
    aVelCapMmS : ARRAY[1..16] OF LREAL;   // 各段允许速度上限输出 [mm/s] / Per-segment velocity cap output [mm/s]
    bPlanned   : BOOL;           // 规划完成，单拍脉冲 [-] / Planning done, single-scan pulse
    bCfgBad    : BOOL;           // 组态非法（锁存） [-] / Illegal configuration, latched
    bError     : BOOL;           // 故障标志（与 bCfgBad 同源，R191） [-] / Error flag
END_VAR
VAR
    _nCount : DINT;              // 钳位后有效段数 [段] / Clamped segment count
    _nDepth : DINT;              // 钳位后前瞻深度（<= 段数-1） [段] / Clamped lookahead depth
    _bGo    : BOOL;              // 本拍规划执行许可（组态合法 ∧ 目标速度正） / Planning permission this scan
    _fVc    : LREAL;             // 单段拐角限速中间量 [mm/s] / Corner speed intermediate
    _fAcc2  : LREAL;             // 回溯/前传累加式中间量 [mm²/s²] / Backward-pass square accumulator
    i       : DINT;              // 段循环索引 / Segment loop index
    _bErrScan: BOOL;             // 当拍错误内部量（超限钳位） / Per-scan error internal
    _bCfgLatch: BOOL;            // 组态非法锁存位（解除沿 = bReset 上升沿） / Latched config fault
    rtReset : R_TRIG;            // 复位沿实例，段 0 无条件调用 / Reset edge instance
END_VAR
VAR CONSTANT
    DL_LVP_NMAX : DINT  := 16;       // 段表定长上限 [段] / Segment table length ceiling
    DL_LVP_ZERO : LREAL := 0.0;      // 判零基准 [无量纲] / Zero base
    DL_LVP_TWO  : LREAL := 2.0;      // 加速距离公式系数 [-] / Kinematics factor two
END_VAR

(* —— 段 0：段数钳位 + 组态闸 + 沿刷新 —— *)
_bErrScan := FALSE;                          // 当拍错预清 / Per-scan error preset
_nCount := UDINT_TO_DINT(nSegCount);         // 段数转 DINT（超界由下步钳位） / Convert count
IF _nCount > DL_LVP_NMAX THEN
    _nCount := DL_LVP_NMAX;                  // 段数钳到定长上限（头注释②） / Clamp count to ceiling
    _bErrScan := TRUE;                       // 记当拍错 / Mark per-scan error
END_IF
IF _nCount < 0 THEN
    _nCount := 0;                            // UDINT 溢出负值兜底 / Overflow fallback
    _bErrScan := TRUE;                       // 记当拍错 / Mark per-scan error
END_IF
_nDepth := UDINT_TO_DINT(nLookahead);        // 前瞻深度转换 / Convert depth
IF _nDepth > (_nCount - 1) THEN
    _nDepth := _nCount - 1;                  // 深度钳到段数-1（回溯窗不出界） / Clamp depth to count-1
END_IF
IF _nDepth < 0 THEN
    _nDepth := 0;                            // 深度非负兜底 / Depth non-negative
END_IF
_bGo := (_nCount >= 1) AND (fVtrajMmS > DL_LVP_ZERO) AND (NOT _bCfgLatch);   // 规划执行许可（段数/速度/组态三闸） / Planning permission
rtReset(CLK := bReset);                      // 复位沿，每拍必调 / Reset edge, every scan

(* —— 段 1：复位沿 —— *)
IF rtReset.Q THEN
    _bCfgLatch := FALSE;                     // 清组态锁存 / Clear cfg latch
END_IF

(* —— 段 2：段几何病校验（fLen/fAccel/fVmax 非正 → 锁存，病态期冻结输出） —— *)
IF _bGo THEN
    FOR i := 1 TO _nCount DO
        IF (aSeg[i].fLenMm <= DL_LVP_ZERO) OR (aSeg[i].fAccelMmS2 <= DL_LVP_ZERO)
           OR (aSeg[i].fVmaxMmS <= DL_LVP_ZERO) THEN
            _bCfgLatch := TRUE;              // 零长度/零加速段：除零隐患前置锁存（头注释③） / Bad segment geometry: latch
        END_IF
    END_FOR
END_IF

(* —— 段 3：三步规划（组态合法期执行；bPlanned 单拍） —— *)
bPlanned := FALSE;                           // 规划脉冲预清 / Planned pulse preset
IF _bGo AND (NOT _bCfgLatch) THEN
    (* 第 1 步：段上限 = MIN(轨迹目标, 段限速, 拐角限速) *)
    FOR i := 1 TO _nCount DO
        aVelCapMmS[i] := fVtrajMmS;          // 目标速度起步 / Start from target speed
        IF aVelCapMmS[i] > aSeg[i].fVmaxMmS THEN
            aVelCapMmS[i] := aSeg[i].fVmaxMmS;   // 段限速钳入 / Clamp to segment ceiling
        END_IF
        _fVc := SQRT(aSeg[i].fAccelMmS2 * aSeg[i].fCornerRad);   // 拐角限速 = √(a×R)（R>=0 保证非负，R6 无负开方） / Corner speed
        IF (aSeg[i].fCornerRad > DL_LVP_ZERO) AND (aVelCapMmS[i] > _fVc) THEN
            aVelCapMmS[i] := _fVc;           // 拐角限速钳入（半径 0 段不限） / Clamp to corner speed
        END_IF
    END_FOR
    (* 第 2 步：自深至浅回溯（减速可达性反推；FOR 定界，等价 WHILE+步数计数防死锁） *)
    FOR i := (_nCount - 1) TO (MAX(_nCount - _nDepth - 1, 1)) BY -1 DO
        _fAcc2 := aVelCapMmS[i + 1] * aVelCapMmS[i + 1] + DL_LVP_TWO * aSeg[i].fAccelMmS2 * aSeg[i].fLenMm;   // 可达平方累加式（减速距离取本段 L[i]，v1.0.1 返修） / Reachable square accumulator, current segment length
        IF _fAcc2 < DL_LVP_ZERO THEN
            _fAcc2 := DL_LVP_ZERO;           // 累加式为负先钳 0 再开方（头注释④） / Clamp negative square
        END_IF
        _fVc := SQRT(_fAcc2);                // 可达速度上限 [mm/s] / Reachable speed
        IF aVelCapMmS[i] > _fVc THEN
            aVelCapMmS[i] := _fVc;           // 回溯降速 / Backward cap
        END_IF
    END_FOR
    (* 第 3 步：前向传播可达上限（加速可达性顺推） *)
    FOR i := 1 TO (_nCount - 1) DO
        _fAcc2 := aVelCapMmS[i] * aVelCapMmS[i] + DL_LVP_TWO * aSeg[i + 1].fAccelMmS2 * aSeg[i + 1].fLenMm;   // 前传平方累加式 / Forward square accumulator
        IF _fAcc2 < DL_LVP_ZERO THEN
            _fAcc2 := DL_LVP_ZERO;           // 累加式为负先钳 0 / Clamp negative square
        END_IF
        _fVc := SQRT(_fAcc2);                // 可达速度上限 / Reachable speed
        IF aVelCapMmS[i + 1] > _fVc THEN
            aVelCapMmS[i + 1] := _fVc;       // 前传降速 / Forward cap
        END_IF
    END_FOR
    bPlanned := TRUE;                        // 规划完成单拍 / Planning done pulse
END_IF

(* —— 段 4：故障出口（名实双出口同源，R191） —— *)
bCfgBad := _bCfgLatch;                       // 组态非法出口 / Cfg fault outlet
bError  := _bCfgLatch OR _bErrScan;          // 故障标志 = 组态锁存 ∨ 当拍超限 / Error flag

END_FUNCTION_BLOCK

(* ---- FB_DL_MoveResumeSeg.st ---- *)
(*==============================================================================
 * 组件名称 (Component)  : FB_DL_MoveResumeSeg
 * 所属子库 (Sublibrary) : DL_Motion
 * 当前版本 (Version)    : 1.0.1
 * 兼容性 (Platform)     : CODESYS 3.5+ / TwinCAT 3 / 汇川 InoProShop / 施耐德 Machine Expert
 *                         仅依赖 Standard.library（R_TRIG），零厂商私有库，
 *                         零轴状态枚举引用（R277：运动层状态属主唯一）
 * 功能描述 (Function)   : 断点续走。运行中按 bSaveCmd 沿快照「起点/目标」对
 *                         （fStartSave/fTargetSave 输出供上层落盘持久化）；
 *                         断电重启后上层把持久化值从 fTargetRst/fStartRst 注入
 *                         并给 bRestore 沿，本件以当前位置计算剩余行程与方向，
 *                         进入续走相：输出方向位与剩余距离，上层以既有运动
 *                         指令件执行；到达容差内 → bResumeDone 单拍并收口。
 * 来源标签 (Origin)     : 自研线（IEC 61131-3 标准语义的道莅防御性实现，clean-room）
 * 分工声明 (Pairing)    : MoveResumeSeg（断点续走，本件）↔ MotionCmdQueue（指令
 *                         排队，既有件）：本件只产出「剩余行程/方向/进度」快照
 *                         与续走判据，不生成运动指令、不排队、不接管轴使能
 *                         （R298 属主边界：续走计算不替代指令编排）。
 * 边界语义 (Boundary)   : ① 进度除零防御：目标 = 起点段长 <= eps → 组态故障
 *                         锁存（零行程快照无续走语义）；
 *                         ② 恢复闸：恢复时位置已在目标容差内 → 直接收口
 *                         bResumeDone，不发续走（防负行程往回走）；
 *                         ③ 剩余距离负值（越过目标）→ 按已到收口，不输出反向
 *                         续走（安全侧）；
 *                         ④ 位置 NaN → 本拍冻结（不派生方向）；
 *                         ⑤ 组态闸：容差 <= 0 / 速度域 → 故障。
 * 输出语义 (Fallback)   : 【R191】bEnable = FALSE → 方向/续走输出强制 FALSE
 *                         （续走是执行建议，失能必须收敛）；eFault 相 → 冻结
 *                         + bError = TRUE。
 * 码位     (Codes)      : 按 R297 范式零 16# 码位硬编码；错误出口 BOOL+ENUM(eCause)，
 *                         码位待主控收口统一派号。
 * 红线自检 (Redline)    : 7 项红线已自检：R1 零全局 ✓｜R2 零物理地址 ✓｜R3 纯 IEC ✓
 *                         R4 除零（段长 eps 闸）/NaN 冻结/组态闸 ✓
 *                         R5 双语同行注释 ✓｜R6 CASE 带 ELSE 兜底迁 eFault ✓
 *                         R7 R_TRIG 段 0 无条件刷新 ✓
 * 验收向量 (Acceptance) : V1 快照 (100, 300)，恢复时位置 220 → 剩余 80，
 *                         bDirPos=TRUE，fProgress=0.6；
 *                         V2 恢复时位置 295（容差 5 内）→ 直接 bResumeDone；
 *                         V3 恢复时位置 310（越目标）→ bResumeDone 不反向；
 *                         V4 快照起点=目标 → eFault 组态锁存。
 * 修订历史 (Revision)   : 2026-11-20  v1.0.0  R49 首版（批 4 · 序号 16）
 *                        2026-11-20  v1.0.1  R51 返修（R50 终审中）：eResume 相方向
 *                        改进入相时锁存（_bDir 不再每拍重派生，R339 方向锁定）；
 *                        越目标（剩余量符号与锁定方向相反）一律按已到收口
 *                        bResumeDone，不输出反向续走（与边界③一致）
 *==============================================================================*)
TYPE E_DL_MrsState :
(
    eIdle    := 0,                           (* 待快照/待恢复 / Idle *)
    eSaved   := 10,                          (* 快照已建立，运行中持续更新进度 / Saved, tracking progress *)
    eResume  := 20,                          (* 续走执行中（方向/剩余距离输出） / Resuming *)
    eDone    := 30,                          (* 续走完成收口保持 / Resume done hold *)
    eFault   := 90                           (* 故障锁存相 / Fault latched phase *)
);
END_TYPE

TYPE E_DL_MrsCause :
(
    eNone       := 0,                        (* 无故障成因 / No cause *)
    eCfgIllegal := 1,                        (* 组态非法：容差越域 / Illegal config *)
    eSegIllegal := 2,                        (* 快照段长非法（起点=目标） / Illegal segment length *)
    ePhaseBad   := 3                         (* 非法相位兜底 / Illegal phase fallback *)
);
END_TYPE

FUNCTION_BLOCK FB_DL_MoveResumeSeg
VAR_INPUT
    fPosNow    : LREAL := 0.0;               (* 当前轴位置（调用方每拍快照传入）[mm] / Current axis position *)
    fTolerance : LREAL := 0.5;               (* 到位容差，域 > 0.0 [mm] / Arrival tolerance *)
    bSaveCmd   : BOOL := FALSE;              (* 快照命令，上升沿以当前段建立快照 [-] / Snapshot command edge *)
    fTargetRst : LREAL := 0.0;               (* 持久化目标位置注入（断电恢复用）[mm] / Restored target position *)
    fStartRst  : LREAL := 0.0;               (* 持久化起点位置注入（预留 reserved：当前正文零引用，起点语义由 fPosNow 实时快照）[mm] / Restored start position, reserved *)
    bRestoreCmd: BOOL := FALSE;              (* 恢复命令，上升沿按注入值续走 [-] / Restore command edge *)
    bAbort     : BOOL := FALSE;              (* 中止电平，TRUE 终止续走回 eIdle（快照保留）[-] / Abort level *)
    bEnable    : BOOL := TRUE;               (* 使能，FALSE 续走输出强制收敛 [-] / Enable *)
    bReset     : BOOL := FALSE;              (* 复位命令，上升沿清全部内部状态 [-] / Reset command *)
END_VAR
VAR_OUTPUT
    bDirPos     : BOOL;                      (* 续走方向位：TRUE 正向 / FALSE 负向 [-] / Resume direction flag *)
    fRemainAbs  : LREAL;                     (* 剩余行程绝对值 [mm] / Remaining distance *)
    fProgress   : LREAL;                     (* 段内完成进度 0..1（快照相实时更新）[-] / Segment progress *)
    bResumeActive : BOOL;                    (* 续走执行中指示 [-] / Resume-active indicator *)
    fTargetSave : LREAL;                     (* 快照目标（供上层持久化落盘）[mm] / Snapshot target for persistence *)
    fStartSave  : LREAL;                     (* 快照起点（供上层持久化落盘）[mm] / Snapshot start for persistence *)
    bResumeDone : BOOL;                      (* 续走完成单拍位 [-] / Resume-done single-scan pulse *)
    eState      : E_DL_MrsState;             (* 状态出口 / State outlet *)
    eCause      : E_DL_MrsCause;             (* 故障成因出口（R190 归因唯一） / Fault cause outlet *)
    bError      : BOOL;                      (* 故障锁存标志 [-] / Fault latch flag *)
END_VAR
VAR
    _eState   : E_DL_MrsState := E_DL_MrsState.eIdle;     (* 内部相位（CASE 唯一写入目标） / Internal phase *)
    _eCause   : E_DL_MrsCause := E_DL_MrsCause.eNone;     (* 故障成因锁存量 / Latched cause *)
    rtSave    : R_TRIG;                     (* 快照沿实例，段 0 无条件调用 / Save edge instance *)
    rtRestore : R_TRIG;                     (* 恢复沿实例，段 0 无条件调用 / Restore edge instance *)
    rtReset   : R_TRIG;                     (* 复位沿实例，段 0 无条件调用 / Reset edge instance *)
    _fTarget  : LREAL;                       (* 目标位置锁存（快照槽）[mm] / Target latch *)
    _fStart   : LREAL;                       (* 起点位置锁存（快照槽）[mm] / Start latch *)
    _fRemain  : LREAL;                       (* 剩余行程派生量 [mm] / Remaining derived *)
    _fSegLen  : LREAL;                       (* 段长派生量 [mm] / Segment length derived *)
    _fProg    : LREAL;                       (* 进度派生量 [-] / Progress derived *)
    _bDir     : BOOL;                        (* 方向锁存量（进入 eResume 相时锁定，越目标不反向，R339）[-] / Direction latch *)
    _bReached : BOOL;                        (* 到位当拍判据 [-] / Reached verdict this scan *)
    _bPosBad  : BOOL;                        (* 位置非有限当拍量 [-] / Non-finite position this scan *)
    _bFault   : BOOL;                        (* 故障锁存位 / Latched fault bit *)
    _bCfgBad  : BOOL;                        (* 组态非法当拍量 / Illegal config this scan *)
END_VAR
VAR CONSTANT
    DL_MRS_EPS : LREAL := 1.0E-9;            (* 段长判零容差 [mm²] / Segment epsilon *)
END_VAR

(* —— 段 0：当拍判据派生 + 沿实例无条件刷新（R228A） —— *)
_bCfgBad := (fTolerance <= 0.0);             (* 组态闸：容差正域（R151 全引脚，单引脚件） / Config gate *)
rtSave(CLK := bSaveCmd);                     (* 快照沿每拍必调 / Save edge every scan *)
rtRestore(CLK := bRestoreCmd);               (* 恢复沿每拍必调 / Restore edge every scan *)
rtReset(CLK := bReset);                      (* 复位沿每拍必调 / Reset edge every scan *)
_bPosBad := (fPosNow <> fPosNow) OR ((fPosNow - fPosNow) <> (fPosNow - fPosNow));   (* 位置 NaN 自反 + Inf 差判 / Non-finite position *)

(* —— 段 1：单拍量预清零（R107） —— *)
bResumeDone := FALSE;                        (* 完成单拍位预清，唯一分支置位 / Done pulse preset *)
_bReached := FALSE;                          (* 到位判据预清 / Reached preset *)
_fRemain := 0.0;                             (* 剩余距离预清（每拍全路径派生，R285） / Remain preset *)
_fProg := 0.0;                               (* 进度预清 / Progress preset *)

(* —— 段 2：复位沿处理（作用域：清故障 + 清快照槽 + 清输出镜像 + 迁 eIdle，R283 逐项声明） —— *)
IF rtReset.Q THEN
    _bFault := FALSE;                        (* 清故障锁存 / Clear fault *)
    _eCause := E_DL_MrsCause.eNone;          (* 清成因 / Clear cause *)
    _fTarget := 0.0;                         (* 清目标槽 / Clear target *)
    _fStart := 0.0;                          (* 清起点槽 / Clear start *)
    fTargetSave := 0.0;                      (* 清快照目标镜像 / Clear mirror *)
    fStartSave := 0.0;                       (* 清快照起点镜像 / Clear mirror *)
    fRemainAbs := 0.0;                       (* 清剩余镜像 / Clear remain *)
    fProgress := 0.0;                        (* 清进度镜像 / Clear progress *)
    bDirPos := FALSE;                        (* 清方向镜像 / Clear direction *)
    _eState := E_DL_MrsState.eIdle;          (* 迁待机相 / Back to idle *)
END_IF

(* —— 段 3：组态闸故障锁存（R45 配对；锁存至复位沿，R189） —— *)
IF _bCfgBad AND NOT _bFault THEN
    _bFault := TRUE;                         (* 锁存故障位 / Latch fault *)
    _eCause := E_DL_MrsCause.eCfgIllegal;    (* 成因：组态非法 / Cause: illegal config *)
    _eState := E_DL_MrsState.eFault;         (* 同步迁故障相 / Migrate to fault *)
END_IF

(* —— 段 4：CASE 主状态机（ELSE 兜底迁 eFault，红线 6） —— *)
CASE _eState OF
    E_DL_MrsState.eIdle:                     (* 待机相 / Idle *)
        IF rtSave.Q AND bEnable AND NOT _bFault AND NOT _bPosBad THEN
            _fStart := fPosNow;              (* 以当前位置建快照起点 / Snapshot start *)
            _fTarget := fTargetRst;          (* 目标取恢复注入口（上层运行中把目标送此口） / Target from injection port *)
            _fSegLen := _fTarget - _fStart;  (* 段长派生 / Segment length *)
            IF ABS(_fSegLen) <= DL_MRS_EPS THEN
                _eCause := E_DL_MrsCause.eSegIllegal;   (* 零行程快照归因（独立分码，R190） / Zero-segment cause *)
                _bFault := TRUE;             (* 故障锁存（R45 配对） / Latch fault *)
                _eState := E_DL_MrsState.eFault;   (* 同步迁故障相 / Migrate to fault *)
            ELSE
                fStartSave := _fStart;       (* 快照起点镜像输出（供上层落盘） / Start mirror *)
                fTargetSave := _fTarget;     (* 快照目标镜像输出 / Target mirror *)
                _eState := E_DL_MrsState.eSaved;   (* 进入快照跟踪 / Enter saved *)
            END_IF
        END_IF
    E_DL_MrsState.eSaved:                    (* 快照跟踪相：实时进度更新 / Saved *)
        IF NOT _bPosBad THEN
            _fSegLen := _fTarget - _fStart;  (* 段长重派生（目标/起点为锁存槽，段长恒定） / Segment length *)
            _fProg := (fPosNow - _fStart) / _fSegLen;   (* 进度派生：除子为段长（快照闸已保证 |段长| > eps），无除零 / Progress, divisor gated *)
            fProgress := _fProg;             (* 进度实时镜像 / Progress mirror *)
        END_IF
        IF rtRestore.Q AND bEnable AND NOT _bFault THEN
            IF NOT _bPosBad THEN
                _fRemain := _fTarget - fPosNow;   (* 剩余行程派生 / Remaining *)
                IF ABS(_fRemain) <= fTolerance THEN
                    bResumeDone := TRUE;     (* 恢复即到位：直接收口（边界②防负行程） / Restore in tolerance: done *)
                    _eState := E_DL_MrsState.eDone;   (* 收口相 / Enter done *)
                ELSE
                    _bDir := (_fRemain > 0.0);   (* 方向锁存：进 eResume 后不再重派生（R339） / Direction latched on entry *)
                    _eState := E_DL_MrsState.eResume;   (* 进入续走 / Enter resume *)
                END_IF
            END_IF
        END_IF
    E_DL_MrsState.eResume:                   (* 续走执行相 / Resume *)
        IF NOT bEnable OR bAbort THEN        (* 失能/中止：输出收敛回待机（快照保留，可再次恢复） / Disable or abort *)
            _eState := E_DL_MrsState.eIdle;  (* 回待机 / Back to idle *)
        ELSIF _bPosBad THEN
            ;                                (* 位置坏值拍：输出冻结保持（边界④），不迁相 / Bad position: freeze *)
        ELSE
            _fRemain := _fTarget - fPosNow;  (* 剩余行程每拍重派生 / Remaining re-derived *)
            IF ABS(_fRemain) <= fTolerance THEN
                bResumeDone := TRUE;         (* 到位收口单拍 / Done pulse *)
                _eState := E_DL_MrsState.eDone;   (* 收口相 / Enter done *)
            ELSIF (_fRemain > 0.0) <> _bDir THEN   (* 越目标：剩余量符号与锁定方向相反（边界③，R339） / Overshoot: sign opposes latched direction *)
                bResumeDone := TRUE;         (* 越目标按已到收口，不反向续走 / Overshoot closes as done, no reversal *)
                _eState := E_DL_MrsState.eDone;   (* 收口相 / Enter done *)
            ELSE
                fRemainAbs := ABS(_fRemain); (* 剩余绝对值镜像 / Remain mirror *)
                bDirPos := _bDir;            (* 方向镜像（取锁存值，不重派生） / Direction mirror from latch *)
            END_IF
        END_IF
    E_DL_MrsState.eDone:                     (* 收口保持相 / Done *)
        IF rtSave.Q AND bEnable AND NOT _bFault AND NOT _bPosBad THEN
            _fStart := fPosNow;              (* 新一轮快照（同 eIdle 建快照语义） / New snapshot *)
            _fTarget := fTargetRst;          (* 目标取注入口 / Target from port *)
            _fSegLen := _fTarget - _fStart;  (* 段长派生 / Segment length *)
            IF ABS(_fSegLen) > DL_MRS_EPS THEN
                fStartSave := _fStart;       (* 快照镜像 / Snapshot mirror *)
                fTargetSave := _fTarget;     (* 快照镜像 / Snapshot mirror *)
                _eState := E_DL_MrsState.eSaved;   (* 回跟踪相 / Back to saved *)
            ELSE
                _eCause := E_DL_MrsCause.eSegIllegal;   (* 零行程归因 / Zero-segment cause *)
                _bFault := TRUE;             (* 故障锁存 / Latch fault *)
                _eState := E_DL_MrsState.eFault;   (* 迁故障相 / To fault *)
            END_IF
        END_IF
    E_DL_MrsState.eFault:                    (* 故障相：冻结保持，仅复位沿出 / Fault *)
        ;                                    (* 锁存回放（R28） / Replay from latch *)
    ELSE                                     (* 非法相位兜底迁安全态 / Illegal phase fallback *)
        _eState := E_DL_MrsState.eFault;     (* 迁故障相 / To fault *)
        _bFault := TRUE;                     (* 同步锁存 / Latch *)
        _eCause := E_DL_MrsCause.ePhaseBad;  (* 成因：非法相位 / Cause: illegal phase *)
END_CASE

(* —— 段 5：出口映射（双门控收敛，R191/R285） —— *)
IF _eState = E_DL_MrsState.eResume AND bEnable AND NOT _bFault AND NOT _bPosBad THEN
    bResumeActive := TRUE;                   (* 续走执行中指示 / Resume-active indicator *)
    bDirPos := _bDir;                        (* 方向出口（续走相每拍已派生） / Direction outlet *)
    fRemainAbs := ABS(_fRemain);             (* 剩余出口 / Remain outlet *)
ELSE
    bResumeActive := FALSE;                  (* 非续走相指示收敛 / Indicator converge *)
    bDirPos := FALSE;                        (* 方向收敛（失能必须收敛语义） / Direction converge *)
END_IF
bError := _bFault;                           (* 故障标志镜像 / Fault flag mirror *)
eState := _eState;                           (* 状态出口 / State outlet *)
eCause := _eCause;                           (* 成因出口 / Cause outlet *)
END_FUNCTION_BLOCK

(* ---- FB_DL_NotchAlignSeq.st ---- *)
(*==============================================================================
 * 组件名称 (Component)  : FB_DL_NotchAlignSeq
 * 所属子库 (Sublibrary) : DL_Motion
 * 当前版本 (Version)    : 1.0.0
 * 兼容性 (Platform)     : CODESYS 3.5 / TwinCAT 3 / 汇川 InoProShop（纯标准元素，零方言）
 * 功能描述 (Function)   : 晶圆缺口对位六相顺控。搜索相等待缺口检出，锁存相用条件加减归
 *                         一角度（禁用取模，负数取余三平台不一致）并算最小转角，微调相
 *                         派发相对转动，复核相按公差判合格，超差在限次内重试，限次用尽
 *                         或单相超时一律锁存故障，不空转。不做缺口视觉识别本身（检出由
 *                         引脚注入）、不做旋转轴回零、不做多片排队。
 *                         说明：I_DL_StepperOpenLoop.MoveRelative 为线性距离语义，本件把
 *                         旋转角度直接按「度」传给距离参数（旋转轴已按 1 mm = 1 ° 标定），
 *                         该标定假设由调用方在轴组态中保证。
 * 溯源 (Origin)         : 道莅 clean-room 防御性实现
 * 本文件内含 (Contains) : TYPE E_DL_NotchState / FUNCTION_BLOCK FB_DL_NotchAlignSeq
 * 依赖 (Depends)        : DL_Device/I_DL_StepperOpenLoop（只调用契约方法与属性）
 * 红线自检 (Redline)    : 无外部全局变量、无硬件地址直引 ｜ 全变量中英双语同行注释
 *                         公差与速度判零防除零 ｜ 角度归一用条件加减（禁取模） ｜ 非有限
 *                         用自反比较 ｜ 相超时定时器与沿实例无条件周期刷新 ｜ 枚举显式赋值
 *                         ｜ 搜索相退出条件 ≥2 条（缺口检出沿 + 前置条件消失/超时） ｜ CASE 含 ELSE
 * 错误码表 (Codes)      : 16#0004_0336 就绪（空闲/完成/无事件）
 *                         16#0004_0337 故障级 旋转轴拒绝微调指令
 *                         16#0004_0338 故障级 组态非法（公差/角速度/相超时/限次出域）
 *                         16#0004_0339 故障级 单相超时（不自动续相，必须复位后重新启动）
 *                         16#0004_033A 故障级 重试次数用尽。本件 5 槽全用、无预留槽，已登记待裁定
 * 修订历史 (Revision)   : 2026-11-17  v1.0.0  首版入库 · R28 · 阶段三批 2
 * 验收向量 (Acceptance) : 正向 当前 10 °、目标 95 °、公差 0.2 °、30 °/s → 微调 +85 °、
 *                         复核偏差 0.05 ° → eDone
 *                         反向 缺口检出恒 FALSE → 超时 16#0004_0339 转 eFault（不空转）；
 *                         公差给 0 → 16#0004_0338；限次 0 且复核超差 → 16#0004_033A
 *============================================================================*)

(*-----------------------------------------------------------------------------
 * 枚举: E_DL_NotchState（归属本功能块，同文件发布，全库唯一定义）
 * 含义: 缺口对位相位，每个成员在 CASE 中有且仅有一个标签。
 *----------------------------------------------------------------------------*)
TYPE E_DL_NotchState :
(
    eIdle      := 0,    // 空闲：等启动沿 / Idle, waiting for the start edge
    eSearching := 10,   // 搜索：等缺口检出或相超时 / Searching, waiting for the notch or the phase timeout
    eLatched   := 20,   // 锁存：本拍算最小转角并派单 / Latched, computing the shortest angle and dispatching
    eTrimming  := 30,   // 微调：等旋转轴就绪 / Trimming, waiting for the rotary axis to be ready
    eVerifying := 40,   // 复核：判偏差是否落公差 / Verifying, checking whether the deviation is inside tolerance
    eDone      := 50,   // 完成：单拍完成脉冲，需新启动沿 / Done, one-scan pulse, a new start edge is required
    eFault     := 99    // 故障：锁存码保持，仅复位沿退出 / Fault, the latch code is held until the reset edge
);
END_TYPE

FUNCTION_BLOCK FB_DL_NotchAlignSeq
VAR_INPUT
    bEnable        : BOOL := FALSE;       // 使能 / Enable
    bStart         : BOOL := FALSE;       // 启动，上升沿启动一次 / Start, the rising edge starts one cycle
    bReset         : BOOL := FALSE;       // 复位，仅故障态生效 / Reset, effective in the fault state only
    bNotchFound    : BOOL := FALSE;       // 缺口检出（引脚注入） / Notch found, injected by the caller
    fThetaNow_deg  : REAL := 0.0;         // 当前转角 [°]，域 0~360 / Present angle in degrees, domain 0 to 360
    fThetaTarget_deg : REAL := 0.0;       // 目标转角 [°]，域 0~360 / Target angle in degrees, domain 0 to 360
    fTolDeg        : REAL := 0.2;         // 复核公差 [°]，域 0.01~1.0 / Verification tolerance in degrees, domain 0.01 to 1.0
    fSpinSpeed_dps : REAL := 30.0;        // 角速度 [°/s]，域 1~180 / Angular speed in degrees per second, domain 1 to 180
    tPhaseMax      : TIME := T#10S;       // 单相超时 [ms]，域 100ms~30s / Per-phase timeout, domain 100 ms to 30 s
    uRetryMax      : UINT := 2;           // 重试上限 [次]，域 0~2 / Retry limit, domain 0 to 2
END_VAR
VAR_IN_OUT
    iAxis          : I_DL_StepperOpenLoop; // 旋转轴开环步进契约引用 [—] / Rotary axis open-loop stepper contract reference
END_VAR
VAR_OUTPUT
    bDone          : BOOL;                // 完成脉冲，单拍有效 / Completion pulse, valid for one scan
    bBusy          : BOOL;                // 顺控进行中 / Sequence running
    bError         : BOOL;                // 故障级标志，仅故障级码置位 / Fault-class flag, set on fault codes only
    fThetaErr_deg  : REAL;                // 最终偏差 [°] / Final deviation in degrees
    uRetryCnt      : UINT;                // 已重试次数 [次] / Retry count
    eState         : E_DL_NotchState;     // 对位相位 [—] / Alignment phase
    eErr           : UDINT;               // 错误码，段位 16#0004_xxxx / Error code in segment 16#0004_xxxx
END_VAR
VAR
    _eState        : E_DL_NotchState := E_DL_NotchState.eIdle; // 当前相位 / Current phase
    _bInit         : BOOL := FALSE;       // 首扫标志，取非判定 / First-scan flag, tested negated
    _bRefOk        : BOOL;                // 契约引用有效标志 / Contract reference valid flag
    _bCfgOk        : BOOL;                // 组态合法标志 / Configuration valid flag
    _bIssueScan    : BOOL;                // 派单当拍标志（本拍不判就绪） / Dispatch scan flag, readiness is not judged in this scan
    _bFaultLatch   : BOOL;                // 故障锁存标志 / Fault latch flag
    _uLatchCode    : UDINT;               // 锁存码载体 / Latch code carrier
    _fDelta        : REAL;                // 本拍最小转角（已归一）[°] / Shortest angle after normalisation in degrees
    _fErrAbs       : REAL;                // 偏差绝对值 [°] / Absolute deviation in degrees
    _rtrigStart    : R_TRIG;              // 启动上升沿 / Rising edge of the start command
    _rtrigReset    : R_TRIG;              // 复位上升沿 / Rising edge of the reset command
    _rtrigNotch    : R_TRIG;              // 缺口检出上升沿 / Rising edge of the notch-found signal
    _tonPhase      : TON;                 // 单相超时计时 / Per-phase timeout timer
END_VAR
VAR CONSTANT
    DL_NA_READY   : UDINT := 16#0004_0336;  // 就绪码 / Ready code
    DL_NA_AXIS_BAD : UDINT := 16#0004_0337; // 故障级轴拒绝码 / Fault code for a rejected axis command
    DL_NA_CFG_BAD : UDINT := 16#0004_0338;  // 故障级组态非法码 / Fault code for bad configuration
    DL_NA_TIMEOUT : UDINT := 16#0004_0339;  // 故障级相超时码 / Fault code for a phase timeout
    DL_NA_RETRY   : UDINT := 16#0004_033A;  // 故障级重试用尽码 / Fault code for exhausted retries
    DL_NA_HALF    : REAL := 180.0;          // 半周角 [°] / Half turn in degrees
    DL_NA_FULL    : REAL := 360.0;          // 全周角 [°] / Full turn in degrees
    DL_NA_TOL_LO  : REAL := 0.01;           // 公差下限 [°] / Tolerance lower bound
    DL_NA_TOL_HI  : REAL := 1.0;            // 公差上限 [°] / Tolerance upper bound
    DL_NA_SPD_LO  : REAL := 1.0;            // 角速度下限 [°/s] / Angular speed lower bound
    DL_NA_SPD_HI  : REAL := 180.0;          // 角速度上限 [°/s] / Angular speed upper bound
END_VAR

// 段 1｜输出与单拍标志预置
bDone := FALSE;                                     // 完成脉冲预清 / Completion pulse pre-cleared
bBusy := FALSE;                                     // 运行标志预清 / Busy flag pre-cleared
bError := FALSE;                                    // 故障标志预清 / Fault flag pre-cleared
eErr := 0;                                          // 错误码预清 / Error code pre-cleared
_bIssueScan := FALSE;                               // 派单当拍标志预清 / Dispatch scan flag pre-cleared
_fErrAbs := 0.0;                                    // 偏差预清 [°] / Deviation pre-cleared

// 段 2｜沿检测无条件周期刷新（严禁置于分支内）
_rtrigStart(CLK := bStart);                         // 启动沿 / Start edge
_rtrigReset(CLK := bReset);                         // 复位沿 / Reset edge
_rtrigNotch(CLK := bNotchFound);                    // 缺口检出沿 / Notch-found edge

// 段 3｜首扫初始化（判据取非，R19）
IF NOT _bInit THEN
    _eState := E_DL_NotchState.eIdle;               // 相位待机起步 / Phase starts idle
    _bInit := TRUE;                                 // 首扫只做一次 / The first scan runs once
END_IF

// 段 4｜引用与组态闸
_bRefOk := (iAxis <> 0);                            // 引用注入判据 / Reference injected flag
_bCfgOk := _bRefOk
        AND NOT ((fTolDeg <> fTolDeg) OR ((fTolDeg - fTolDeg) <> (fTolDeg - fTolDeg)))
        AND (fTolDeg >= DL_NA_TOL_LO) AND (fTolDeg <= DL_NA_TOL_HI)
        AND NOT ((fSpinSpeed_dps <> fSpinSpeed_dps) OR ((fSpinSpeed_dps - fSpinSpeed_dps) <> (fSpinSpeed_dps - fSpinSpeed_dps)))
        AND (fSpinSpeed_dps >= DL_NA_SPD_LO) AND (fSpinSpeed_dps <= DL_NA_SPD_HI)
        AND (tPhaseMax >= T#100MS) AND (tPhaseMax <= T#30S)
        AND (uRetryMax <= 2);

// 段 5｜相超时定时器无条件周期刷新（搜索/锁存/微调/复核四相计时）
_tonPhase(IN := (_eState = E_DL_NotchState.eSearching) OR (_eState = E_DL_NotchState.eLatched)
            OR (_eState = E_DL_NotchState.eTrimming) OR (_eState = E_DL_NotchState.eVerifying),
          PT := tPhaseMax);

// 段 6｜角度归一（条件加减，禁取模；输入域 0~360 故单次修正即落 (-180, 180]）
_fDelta := fThetaTarget_deg - fThetaNow_deg;        // 原始角差 [°] / Raw angle difference
IF _fDelta > DL_NA_HALF THEN
    _fDelta := _fDelta - DL_NA_FULL;                // 大于半周：减一周 [°] / Above half a turn, subtract one turn
END_IF
IF _fDelta <= (0.0 - DL_NA_HALF) THEN
    _fDelta := _fDelta + DL_NA_FULL;                // 小于负半周：加一周 [°] / Below minus half a turn, add one turn
END_IF
_fErrAbs := ABS(_fDelta);                           // 偏差绝对值 [°] / Absolute deviation
fThetaErr_deg := _fErrAbs;                          // 偏差出口 [°] / Deviation output

// 段 7｜失能闸
IF NOT bEnable THEN
    _eState := E_DL_NotchState.eIdle;               // 相位回空闲 / Phase back to idle
    eErr := DL_NA_READY;                            // 失能为正常停机 / Disable is a normal stop
END_IF

// 段 8｜对位状态机（ENUM + CASE + ELSE 兜底）
IF bEnable THEN
    CASE _eState OF

        E_DL_NotchState.eIdle:                      // 空闲：等启动沿，先做组态闸
            IF _rtrigStart.Q THEN
                _bFaultLatch := FALSE;              // 启动沿为锁存解除路径 / The start edge releases the latch
                _uLatchCode := 0;                   // 锁存码清 / Latch code cleared
                uRetryCnt := 0;                     // 重试计数清 [次] / Retry count cleared
                IF NOT _bCfgOk THEN
                    eErr := DL_NA_CFG_BAD;          // 故障级：组态非法 / Fault, bad configuration
                    _uLatchCode := DL_NA_CFG_BAD;
                    _bFaultLatch := TRUE;
                    bError := TRUE;
                    _eState := E_DL_NotchState.eFault;
                ELSE
                    _eState := E_DL_NotchState.eSearching;   // 进入搜索相 / Enter the searching phase
                END_IF
            END_IF

        E_DL_NotchState.eSearching:                 // 搜索：退出条件两条（检出沿 / 超时）
            bBusy := TRUE;
            IF _rtrigNotch.Q THEN
                _eState := E_DL_NotchState.eLatched;         // 条件一：缺口检出 / Condition one, the notch was found
            ELSIF _tonPhase.Q THEN
                eErr := DL_NA_TIMEOUT;                       // 故障级：搜索相超时，不空转 / Fault, searching timed out
                _uLatchCode := DL_NA_TIMEOUT;
                _bFaultLatch := TRUE;
                bError := TRUE;
                bBusy := FALSE;
                _eState := E_DL_NotchState.eFault;           // 条件二：前置条件消失（超时）/ Condition two, the precondition vanished
            END_IF

        E_DL_NotchState.eLatched:                   // 锁存：偏差已在公差内直接复核，否则派单微调
            bBusy := TRUE;
            IF _fErrAbs <= fTolDeg THEN
                _eState := E_DL_NotchState.eVerifying;      // 已到位：直接复核 / Already aligned, go verifying
            ELSIF ABS(_fDelta) > (DL_NA_HALF + DL_NA_TOL_HI) THEN
                eErr := DL_NA_CFG_BAD;                      // 故障级：归一失配（角度输入出域）/ Fault, normalisation mismatch
                _uLatchCode := DL_NA_CFG_BAD;
                _bFaultLatch := TRUE;
                bError := TRUE;
                bBusy := FALSE;
                _eState := E_DL_NotchState.eFault;
            ELSE
                IF iAxis.MoveRelative(_fDelta, fSpinSpeed_dps) THEN
                    _bIssueScan := TRUE;                    // 派单当拍不判就绪 / Readiness is not judged in the dispatch scan
                    _eState := E_DL_NotchState.eTrimming;   // 进入微调相 / Enter the trimming phase
                ELSE
                    eErr := DL_NA_AXIS_BAD;                 // 故障级：轴拒绝指令 / Fault, the axis rejected the command
                    _uLatchCode := DL_NA_AXIS_BAD;
                    _bFaultLatch := TRUE;
                    bError := TRUE;
                    bBusy := FALSE;
                    _eState := E_DL_NotchState.eFault;
                END_IF
            END_IF

        E_DL_NotchState.eTrimming:                  // 微调：等轴就绪或超时
            bBusy := TRUE;
            IF _bIssueScan THEN
                _bIssueScan := FALSE;                       // 派单拍已过 / The dispatch scan has passed
            ELSIF iAxis.bReady THEN
                _eState := E_DL_NotchState.eVerifying;      // 轴就绪：复核 / Axis ready, go verifying
            ELSIF _tonPhase.Q THEN
                eErr := DL_NA_TIMEOUT;                      // 故障级：微调相超时 / Fault, trimming timed out
                _uLatchCode := DL_NA_TIMEOUT;
                _bFaultLatch := TRUE;
                bError := TRUE;
                bBusy := FALSE;
                _eState := E_DL_NotchState.eFault;
            END_IF

        E_DL_NotchState.eVerifying:                 // 复核：合格即完成，超差在限次内重试
            bBusy := TRUE;
            IF _bIssueScan THEN
                _bIssueScan := FALSE;
            ELSIF _tonPhase.Q THEN
                eErr := DL_NA_TIMEOUT;                      // 故障级：复核相超时 / Fault, verifying timed out
                _uLatchCode := DL_NA_TIMEOUT;
                _bFaultLatch := TRUE;
                bError := TRUE;
                bBusy := FALSE;
                _eState := E_DL_NotchState.eFault;
            ELSE
                IF _fErrAbs <= fTolDeg THEN
                    _eState := E_DL_NotchState.eDone;       // 合格 / Accepted
                ELSIF uRetryCnt >= uRetryMax THEN
                    eErr := DL_NA_RETRY;                    // 故障级：重试次数用尽 / Fault, retries exhausted
                    _uLatchCode := DL_NA_RETRY;
                    _bFaultLatch := TRUE;
                    bError := TRUE;
                    bBusy := FALSE;
                    _eState := E_DL_NotchState.eFault;
                ELSE
                    uRetryCnt := uRetryCnt + 1;             // 重试计数 +1 [次] / Retry count incremented
                    _eState := E_DL_NotchState.eSearching;  // 重新搜索 / Search again
                END_IF
            END_IF

        E_DL_NotchState.eDone:                      // 完成：单拍脉冲（下一拍段 1 预清即自清，R24 三律）
            bDone := TRUE;
            bBusy := FALSE;
            eErr := DL_NA_READY;                    // 就绪/完成码 / Ready or completion code
            _eState := E_DL_NotchState.eIdle;       // 需新启动沿重启 / A new start edge is required

        E_DL_NotchState.eFault:                     // 故障：锁存码保持，仅复位沿退出
            bBusy := FALSE;
            eErr := _uLatchCode;                    // 锁存码回放 / Replay the latch code
            bError := TRUE;
            IF _rtrigReset.Q THEN
                IF _bRefOk THEN
                    iAxis.Reset();                  // 轴故障复位 / Axis fault reset
                END_IF
                _bFaultLatch := FALSE;              // 锁存解除 / Latch released
                _uLatchCode := 0;                   // 锁存码清 / Latch code cleared
                uRetryCnt := 0;                     // 重试计数清 [次] / Retry count cleared
                eErr := DL_NA_READY;                // 复位后回就绪码 / Ready code after the reset
                bError := FALSE;
                _eState := E_DL_NotchState.eIdle;   // 回空闲需新启动沿 / Back to idle, a new start edge is required
            END_IF

        ELSE
            // 非法状态兜底（故障级）
            eErr := DL_NA_CFG_BAD;                  // 故障级：非法相位 / Fault, illegal phase
            _uLatchCode := DL_NA_CFG_BAD;
            _bFaultLatch := TRUE;
            bError := TRUE;
            bBusy := FALSE;
            _eState := E_DL_NotchState.eFault;

    END_CASE
END_IF

eState := _eState;                                  // 相位出口镜像 / Phase mirrored to the output pin
END_FUNCTION_BLOCK

(* ---- FB_DL_PathCornerBlend.st ---- *)
(*
  ==================================================================
  组件名 Component  : FB_DL_PathCornerBlend
  分类   Category   : DL_Motion
  复杂度 Complexity  : 中
  版本   Version    : 1.0.0
  功能   Purpose    : 路径拐角圆滑过渡解算。给定方向改变角 fCornerAngDeg 与
                      拐角半径 fBlendR：切点距 fTanLen = R / tan(θ/2)（θ 为
                      方向改变角）；弦高误差 fChordErr = R·(1−cos(θ/2))；误
                      差带超限时按 Rmax = TolErr/(1−cos(θ/2)) 自动回夹半径并
                      置 bClamped；单调性自检：切点距不得超过两相邻段长一半
                      （与 FC_DL_LookaheadVelPlanner 速度前瞻分工互引）。
  来源   Source     : T1-6-plcopen（PLCopen 运动公开语义）
  溯源   Origin     : 圆弧过渡切点/弦高为公开几何语义，clean-room 自研实现，
                      未复制 PLCopen 或任何厂商私有库源码。
  平台   Platform   : 纯 IEC 61131-3，CODESYS / TwinCAT / InoProShop 通用
  分工声明 Split     : 与 FC_DL_LookaheadVelPlanner 分工——后者做段间速度前
                      瞻，本件做拐角几何过渡解算。
  作者   Author     : 道莅代码库 · PLC 编程专家（R59）
  ------------------------------------------------------------------
  边界 Boundary     :
                      一 非有限入参闸（自反双判据，五参数全覆盖）：命中置
                         bError，输出安全侧零（四段式 R45）；
                      二 角度域闸：方向改变角钳入 [1, 179] 度（信息级
                         bClamped），防 tan/cos 小角爆炸与退化；
                      三 除零闸：tan(θ/2) ≤ eps 判退化置 bError；半径自动
                         回夹除式 (1−cos(θ/2)) > eps 由角度域闸保证并显式
                         再闸一层；
                      四 单调性自检：fTanLen > 0.5·min(段A, 段B) 置 bTooLong
                         （交接约束，信息级非故障）；
                      五 无全局变量、无外部变量声明、无物理地址寻址。
  修订记录 Revision  :
    2026-11-21  v1.0.0  R59 首版（批 2 · 序号 10）
  ==================================================================
*)

FUNCTION_BLOCK FB_DL_PathCornerBlend
VAR_INPUT
    fCornerAngDeg : LREAL := 90.0;  // 方向改变角 [度]，域 [1,179] / the direction change angle [degree]
    fBlendR       : LREAL := 10.0;  // 拐角半径 [毫米] / the corner radius [millimeter]
    fTolErr       : LREAL := 0.1;   // 弦高误差带 [毫米] / the chord error band [millimeter]
    fSegLenA      : LREAL := 100.0; // 前段长 [毫米] / the former segment length [millimeter]
    fSegLenB      : LREAL := 100.0; // 后段长 [毫米] / the latter segment length [millimeter]
    bCalc         : BOOL := TRUE;   // 解算使能，失能输出安全侧零 [-] / the calc enable, disabling zeroes the outlets
END_VAR
VAR_OUTPUT
    fTanLen   : LREAL := 0.0; // 切点距拐角距离（两腿对称）[毫米] / the tangent distance from the corner [millimeter]
    fChordErr : LREAL := 0.0; // 弦高误差 [毫米] / the chord sagitta error [millimeter]
    bValid    : BOOL := FALSE; // 解算受理且可用 [-] / the solved and usable flag
    bErrBand  : BOOL := FALSE; // 弦高超误差带（信息级）[-] / the chord beyond the band, informational
    bTooLong  : BOOL := FALSE; // 切点距超段长一半（单调性自检，信息级）[-] / the tangent beyond the half segment, informational
    bClamped  : BOOL := FALSE; // 半径自动回夹发生（信息级）[-] / the radius auto clamp happened, informational
    bError    : BOOL := FALSE; // 故障标志（非有限或退化角）[-] / the fault flag
END_VAR
VAR CONSTANT
    DL_PCB_EPS     : LREAL := 1.0E-9;             // 退化阈值 [无量纲] / the degenerate threshold
    DL_PCB_ANGMIN  : LREAL := 1.0;                // 角度域下界 [度] / the angle floor
    DL_PCB_ANGMAX  : LREAL := 179.0;              // 角度域上界 [度] / the angle ceiling
    DL_PCB_DEG2RAD : LREAL := 0.0174532925199433; // 度到弧度系数 [弧度每度] / the degree to radian factor
END_VAR
VAR
    lrAng   : LREAL; // 角度工作量（钳后）[度] / the clamped angle work value
    lrHalf  : LREAL; // 半角工作量 [弧度] / the half angle in radian
    lrTanH  : LREAL; // 半角正切工作量 [无量纲] / the half angle tangent
    lrCosH  : LREAL; // 半角余弦工作量 [无量纲] / the half angle cosine
    lrR     : LREAL; // 半径工作量（可回夹）[毫米] / the radius work value, clampable
    lrRmax  : LREAL; // 误差带反算半径上界 [毫米] / the radius bound from the error band
    lrSegMin: LREAL; // 两段较短者 [毫米] / the shorter of the two segments
    bFin    : BOOL;  // 入参有限工作量 [-] / the input finiteness work flag
END_VAR

// 段 1｜输出预置与失能安全侧（四段式，R45）/ segment 1, the preset and the disabled safe side
fTanLen := 0.0; // 切点距预置零 / preset the tangent zero
fChordErr := 0.0; // 弦高预置零 / preset the chord zero
bValid := FALSE; // 有效预置假 / preset the valid false
bErrBand := FALSE; // 超带预置假 / preset the band flag false
bTooLong := FALSE; // 超长预置假 / preset the too long false
bClamped := FALSE; // 回夹预置假 / preset the clamp false
bError := FALSE; // 故障预置假 / preset the fault false
IF NOT bCalc THEN // 失能：输出保持安全侧零 / disabled, keep the safe zero
    RETURN; // 早退 / return early
END_IF

// 段 2｜非有限入参闸（五参数自反双判据全覆盖，R79）/ segment 2, the non finite gate
bFin := (fCornerAngDeg = fCornerAngDeg) AND ((fCornerAngDeg - fCornerAngDeg) = (fCornerAngDeg - fCornerAngDeg)) // 角度有限 / the angle finite
    AND (fBlendR = fBlendR) AND ((fBlendR - fBlendR) = (fBlendR - fBlendR)) // 半径有限 / the radius finite
    AND (fTolErr = fTolErr) AND ((fTolErr - fTolErr) = (fTolErr - fTolErr)) // 误差带有限 / the band finite
    AND (fSegLenA = fSegLenA) AND ((fSegLenA - fSegLenA) = (fSegLenA - fSegLenA)) // 前段有限 / the former finite
    AND (fSegLenB = fSegLenB) AND ((fSegLenB - fSegLenB) = (fSegLenB - fSegLenB)); // 后段有限 / the latter finite
IF NOT bFin THEN // 非有限命中 / a non finite hit
    bError := TRUE; // 置故障（本库纪律②不静默吞）/ raise the fault
    RETURN; // 早退 / return early
END_IF

// 段 3｜角度域钳制与三角量解算（除零前置闸，边界二三）/ segment 3, the angle clamp and the trigonometry
lrAng := fCornerAngDeg; // 装角度 / load the angle
IF lrAng < DL_PCB_ANGMIN THEN // 小角下钳（防 tan 爆炸）/ clamp the small angle
    lrAng := DL_PCB_ANGMIN; // 夹到下界 / clamp to the floor
    bClamped := TRUE; // 信息级 / informational
ELSIF lrAng > DL_PCB_ANGMAX THEN // 大角上钳（防退化）/ clamp the large angle
    lrAng := DL_PCB_ANGMAX; // 夹到上界 / clamp to the ceiling
    bClamped := TRUE; // 信息级 / informational
END_IF
lrHalf := lrAng * 0.5 * DL_PCB_DEG2RAD; // 半角弧度 / the half angle radian
lrTanH := TAN(lrHalf); // 半角正切 / the tangent
lrCosH := COS(lrHalf); // 半角余弦 / the cosine
IF ABS(lrTanH) < DL_PCB_EPS THEN // 退化角闸（切点距无界）/ the degenerate angle gate
    bError := TRUE; // 置故障 / raise the fault
    RETURN; // 早退 / return early
END_IF
lrR := ABS(fBlendR); // 半径取绝对值 / the radius absolute
fTanLen := lrR / lrTanH; // 切点距（除子已闸）/ the tangent distance, divided by the gated tan
fChordErr := lrR * (1.0 - lrCosH); // 弦高误差 / the chord error

// 段 4｜误差带回夹与单调性自检（单点回夹防互相覆盖，边界三四）/ segment 4, the band clamp and the monotonic check
bErrBand := fChordErr > fTolErr; // 超带判定 / the band verdict
IF bErrBand THEN // 超带：反算半径上界回夹 / beyond the band, recompute the radius bound
    IF (1.0 - lrCosH) > DL_PCB_EPS THEN // 除零再闸（角度域已保证，纵深）/ the divide gate, defense in depth
        lrRmax := fTolErr / (1.0 - lrCosH); // 半径上界 [毫米] / the radius bound
        fTanLen := lrRmax / lrTanH; // 回夹后切点距（除子已闸）/ the clamped tangent
        fChordErr := fTolErr; // 弦高回到带上（单点回夹口径）/ the chord to the band
        bClamped := TRUE; // 信息级回夹 / the informational clamp
    ELSE // 反算除子退化（不可达分支兜底）/ the unreachable fallback
        bError := TRUE; // 置故障 / raise the fault
        RETURN; // 早退 / return early
    END_IF
END_IF
lrSegMin := fSegLenA; // 取较短段 / take the shorter segment
IF fSegLenB < lrSegMin THEN // 后段更短 / the latter shorter
    lrSegMin := fSegLenB; // 换取 / take it
END_IF
bTooLong := fTanLen > (0.5 * lrSegMin); // 单调性自检（切点距 ≤ 半段长）/ the monotonic check
bValid := TRUE; // 解算可用 / the solve usable
END_FUNCTION_BLOCK
